(* IEC 61131-3 sources: daoli-st-library/DL_Device (part 26) *)

(* ---- FB_DL_MfcFlowCtrl.st ---- *)
(*==============================================================================
 * 组件名称 (Component)  : FB_DL_MfcFlowCtrl
 * 所属子库 (Sublibrary) : DL_Device
 * 当前版本 (Version)    : 1.0.1
 * 兼容性 (Platform)     : CODESYS 3.5 / TwinCAT 3 / 汇川 InoProShop / Machine Expert
 *                         仅依赖纯 IEC 61131-3 标准元素，零厂商方言
 * 功能描述 (Function)   : MFC 设定-回读校验：新设定上升沿启动跟踪窗，窗内峰值
 *                         对设定+超调阈判超调；回读持续 tStable 在容差窗内判
 *                         入容差；跟踪窗超时（tStable x 5）未入窗 → 稳定超时故障。
 *                         设定 0 视为关断不校验；回读 NaN/越量程判无效冻结。
 * 溯源 (Origin)         : 道莅 clean-room 防御性实现
 * 本文件内含 (Contains) : TYPE E_DL_MfcState / TYPE E_DL_MfcErr /
 *                         FUNCTION_BLOCK FB_DL_MfcFlowCtrl
 * 依赖 (Depends)        : DL_MathData/FC_DL_TimeToDintMs、DL_MathData/FC_DL_TimeScaleSat
 * 红线自检 (Redline)    : 无外部全局变量、无硬件地址直引 ｜ 全变量中英双语同行注释
 *                         防除零 + 参数下限钳制 + 非有限值防御 ｜ 枚举成员全部显式赋值
 *                         TON/沿检测实例每周期无条件调用（仅 IN 条件化）｜
 *                         跟踪窗状态机 CASE 含 ELSE 兜底 ｜ 峰值检测用比较禁浮点判等
 * 错误码表 (Codes)      : 16#0003_0398 就绪
 *                         16#0003_0399 校验通过
 *                         16#0003_039A 信息级 超调检出（不阻断判据）
 *                         16#0003_039B 故障级 稳定超时
 *                         16#0003_039C 故障级 回读无效（冻结判定）
 * 修订历史 (Revision)   : 2026-11-17  v1.0.0  首版入库 · R27 · 阶段三批 2
 *                         2026-11-17  v1.0.1  R27 终审修复（对外引脚零变更）：超调峰值改为
 *                         「首次入窗后才累积、初值取设定」。原实现 fPeakSlm 初值取当前回读，
 *                         降设定（如 20→10 slm）时回读 20 立即满足 20−10 > 超调阈，
 *                         每次下调设定必误报 039A 超调；改为入窗锁存后，仅真实向上超调计入。
 * 验收向量 (Acceptance) : 设定 10 slm 容差 2%FS 超调阈 5%FS：回读峰值 11.0 slm
 *                         → 超调 10%FS → 039A；回读持续 5 s 在 9.8~10.2 → 0399；
 *                         回读 8 slm 持续 25 s → 039B
 *============================================================================*)

(*-----------------------------------------------------------------------------
 * 枚举: E_DL_MfcState（归属 DL_Device，跟踪窗状态机状态）
 *----------------------------------------------------------------------------*)
TYPE E_DL_MfcState :
(
    eIdle    := 0,    // 就绪待新设定 / Idle, waiting for a new setpoint
    eTrack   := 10,   // 跟踪窗：峰值检测与入窗监视 / Tracking window, peak and entry watch
    eStable  := 20,   // 稳定窗：持续容差内计时 / Stable window, dwell timing
    eDone    := 30,   // 校验通过（可被新设定重开）/ Verification passed
    eTimeout := 40,   // 稳定超时故障 / Stable timeout fault
    eFault   := 99    // 回读无效兜底态 / Readback-invalid fallback
);
END_TYPE

(*-----------------------------------------------------------------------------
 * 枚举: E_DL_MfcErr（归属 DL_Device，与 FB_DL_MfcFlowCtrl 同文件）
 *----------------------------------------------------------------------------*)
TYPE E_DL_MfcErr :
(
    eReady      := 16#0003_0398,   // 就绪 / Ready
    ePass       := 16#0003_0399,   // 校验通过 / Verification passed
    eOvershoot  := 16#0003_039A,   // 信息级：超调检出 / Info: overshoot detected
    eStableTmo  := 16#0003_039B,   // 故障级：稳定超时 / Fault: stable timeout
    eReadbackBad:= 16#0003_039C    // 故障级：回读无效 / Fault: readback invalid
);
END_TYPE

(*==============================================================================
 * 功能块: FB_DL_MfcFlowCtrl
 * 调用约定: 每个扫描周期无条件调用一次；tSampleTime 注入真实任务间隔。
 *============================================================================*)
FUNCTION_BLOCK FB_DL_MfcFlowCtrl
VAR_INPUT
    fSetpointSlm   : REAL;            // 设定流量 [标准升每分钟]，有效域 0~满量程 / Setpoint flow [slm]
    fReadbackSlm   : REAL;            // 回读流量 [标准升每分钟] / Readback flow [slm]
    fScaleMaxSlm   : REAL;            // MFC 满量程 [标准升每分钟]，须 > 0 / MFC full scale [slm]
    fTolPct        : REAL := 2.0;     // 容差 [%FS]，默认 2，下限钳 0.5 / Tolerance [percent of FS]
    fOvershootPct  : REAL := 5.0;     // 超调判据 [%FS]，默认 5，下限钳 0.5 / Overshoot criterion [percent of FS]
    tStable        : TIME := T#5S;    // 稳定窗时长 [秒] / Stable window duration [s]
    bNewSp         : BOOL;            // 新设定触发（上升沿）/ New setpoint trigger, rising edge
    tSampleTime    : TIME := T#100MS; // 采样周期，调用方注入 / Sample period, caller-injected
END_VAR
VAR_OUTPUT
    bInTol         : BOOL;            // 入容差标志 / Within-tolerance flag
    bOvershoot     : BOOL;            // 超调检出标志 / Overshoot detected flag
    tSettleMs      : UDINT;           // 实测稳定时间 [毫秒] / Measured settle time [ms]
    eError         : E_DL_MfcErr;     // 错误码 / Error code
    eState         : E_DL_MfcState;   // 跟踪窗状态机当前状态 / Tracking window state
END_VAR
VAR
    fbNewSpTrig    : R_TRIG;          // 新设定上升沿实例（无条件调用）/ New setpoint edge instance
    fbTonStable    : TON;             // 稳定窗计时器（无条件调用）/ Stable window timer
    fbTonWindow    : TON;             // 跟踪窗超时计时器（无条件调用）/ Tracking window timeout timer
    fPeakSlm       : REAL;            // 跟踪窗内回读峰值 [标准升每分钟] / Readback peak in window [slm]
    fTolAbs        : REAL;            // 容差绝对值 [标准升每分钟] / Tolerance in absolute flow [slm]
    fOverAbs       : REAL;            // 超调阈绝对值 [标准升每分钟] / Overshoot threshold in absolute flow [slm]
    fSpUse         : REAL;            // 生效设定（NaN 兜底）[标准升每分钟] / Effective setpoint [slm]
    fScaleUse      : REAL;            // 生效满量程（NaN 兜底）[标准升每分钟] / Effective full scale [slm]
    bReadOk        : BOOL;            // 回读有效性判据 / Readback validity predicate
    uMsErr         : UDINT;           // 委托时间换算错误码（0 = 无错）/ Delegate time-conversion error id
    bInWin         : BOOL;            // 回读在容差窗内（瞬时）/ Readback within window, instantaneous
    bReached       : BOOL;            // 本窗内首次入窗锁存（v1.0.1：峰值仅此后计入）/ First-in-window latch, peak counted afterwards
END_VAR
VAR CONSTANT
    DL_MFC_TOL_MIN    : REAL := 0.5;     // 容差下限 [%FS] / Tolerance lower bound [percent FS]
    DL_MFC_OVER_MIN   : REAL := 0.5;     // 超调阈下限 [%FS] / Overshoot lower bound [percent FS]
    DL_MFC_PCT        : REAL := 100.0;   // 百分数系数 [百分数] / Percent factor
    DL_MFC_WINDOW_K   : INT  := 5;       // 跟踪窗超时倍率（tStable x 5）/ Tracking window timeout multiplier
    DL_MFC_INF_MAX    : REAL := 1.0E30;  // 非有限值判定幅值上限 / Magnitude bound for finite-value check
    DL_MFC_ZERO       : REAL := 0.0;     // 零值常量，避免裸字面量 / Zero constant
    DL_MFC_MS_CAP     : UDINT := 16#FFFF_FFFE;   // 稳定时间输出饱和值 [毫秒] / Settle time saturation [ms]
END_VAR

(*------------------------------------------------------------------------------
 * 段 1｜沿检测与 TON 实例每周期无条件调用（仅 IN 条件化）
 *----------------------------------------------------------------------------*)
fbNewSpTrig(CLK := bNewSp);                           // 新设定沿检测无条件刷新 / new setpoint edge refreshed unconditionally
fbTonStable(IN := (eState = E_DL_MfcState.eStable) AND bInWin, PT := tStable);        // 稳定窗计时 / stable dwell timing
fbTonWindow(IN := (eState = E_DL_MfcState.eTrack), PT := FC_DL_TimeScaleSat(tIn := tStable, nScale := DL_MFC_WINDOW_K));   // 跟踪窗超时计时（tStable x 5，委托换算）/ tracking window timing via delegate

(*------------------------------------------------------------------------------
 * 段 2｜参数防御：满量程/设定 NaN 兜底，容差与超调下限钳 0.5 %FS
 *----------------------------------------------------------------------------*)
fScaleUse := fScaleMaxSlm;                            // 满量程工作副本 / full-scale working copy
IF (fScaleUse <> fScaleUse) OR (fScaleUse <= DL_MFC_ZERO) OR (fScaleUse > DL_MFC_INF_MAX) THEN
    fScaleUse := 100.0;                               // 满量程非法按 100 slm 兜底 / illegal full scale falls back to 100 slm
END_IF
fSpUse := fSetpointSlm;                               // 设定工作副本 / setpoint working copy
IF (fSpUse <> fSpUse) OR (ABS(fSpUse) > DL_MFC_INF_MAX) THEN
    fSpUse := DL_MFC_ZERO;                            // 设定非有限按 0（关断语义）/ non-finite setpoint treated as zero
END_IF
IF fTolPct < DL_MFC_TOL_MIN THEN
    fTolAbs := fScaleUse * DL_MFC_TOL_MIN / DL_MFC_PCT;   // 容差下限钳制 [标准升每分钟] / tolerance floored [slm]
ELSIF fTolPct > DL_MFC_PCT THEN
    fTolAbs := fScaleUse;                             // 容差上限钳制（满量程封顶）/ tolerance capped at FS
ELSE
    fTolAbs := fScaleUse * fTolPct / DL_MFC_PCT;      // 容差换算 [标准升每分钟] / tolerance computed [slm]
END_IF
IF fOvershootPct < DL_MFC_OVER_MIN THEN
    fOverAbs := fScaleUse * DL_MFC_OVER_MIN / DL_MFC_PCT;   // 超调阈下限钳制 / overshoot floored
ELSIF fOvershootPct > DL_MFC_PCT THEN
    fOverAbs := fScaleUse;                            // 超调阈上限钳制 / overshoot capped at FS
ELSE
    fOverAbs := fScaleUse * fOvershootPct / DL_MFC_PCT;   // 超调阈换算 / overshoot computed
END_IF

(*------------------------------------------------------------------------------
 * 段 3｜回读有效性判据：NaN/越量程/负值判无效（bReadOk 为 FALSE 时冻结判定）
 *----------------------------------------------------------------------------*)
bReadOk := (fReadbackSlm = fReadbackSlm)                      // 自反判 NaN / NaN self-reflexive test
        AND (ABS(fReadbackSlm) <= DL_MFC_INF_MAX)             // 溢出判 / overflow test
        AND (fReadbackSlm >= DL_MFC_ZERO)                     // 负流量无效 / negative flow invalid
        AND (fReadbackSlm <= fScaleUse * 1.5);                // 越量程 150% 判无效 / over-range 150 percent invalid

(*------------------------------------------------------------------------------
 * 段 4｜瞬时入窗判据：|回读 - 设定| <= 容差（比较判据，禁浮点判等）
 *----------------------------------------------------------------------------*)
bInWin := bReadOk AND (ABS(fReadbackSlm - fSpUse) <= fTolAbs);   // 瞬时入窗 / instantaneous in-window
IF bInWin THEN
    bReached := TRUE;                                 // v1.0.1：首次入窗锁存，此后峰值才计 / latch on first entry, peak counted after
END_IF
bInTol := bInWin AND fbTonStable.Q AND (eState <> E_DL_MfcState.eIdle);   // 入容差 = 瞬时 + 持续达时 / in-tol combined

(*------------------------------------------------------------------------------
 * 段 5｜新设定上升沿：重开跟踪窗（设定 0 关断不校验，直回就绪）
 *----------------------------------------------------------------------------*)
IF fbNewSpTrig.Q THEN
    IF (fSpUse <= DL_MFC_ZERO) OR (NOT bReadOk) THEN
        eState := E_DL_MfcState.eIdle;                // 设定 0 或回读无效：不启动校验 / zero setpoint or bad readback: no verify
    ELSE
        eState := E_DL_MfcState.eTrack;               // 启动跟踪窗 / start tracking window
        fPeakSlm := fSpUse;                           // v1.0.1：峰值初值取设定而非回读 / peak preset to setpoint, not readback
        bReached := FALSE;                            // v1.0.1：首次入窗锁存清零 / first-entry latch cleared
        bOvershoot := FALSE;                          // 超调标志清零 / overshoot flag cleared
        tSettleMs := 0;                               // 稳定时间清零 / settle time cleared
    END_IF
END_IF

(*------------------------------------------------------------------------------
 * 段 6｜跟踪窗状态机：CASE 含 ELSE 兜底
 *----------------------------------------------------------------------------*)
CASE eState OF

    E_DL_MfcState.eIdle:
        bInTol := FALSE;                              // 就绪态无入容差 / no in-tol in idle
        bOvershoot := FALSE;                          // 就绪态无超调 / no overshoot in idle
        tSettleMs := 0;                               // 稳定时间清零 / settle time cleared
        eError := E_DL_MfcErr.eReady;                 // 码 0398 / code ready

    E_DL_MfcState.eTrack:
        IF bReadOk AND bReached THEN
            IF fReadbackSlm > fPeakSlm THEN
                fPeakSlm := fReadbackSlm;             // 峰值更新（仅首次入窗后计入，禁浮点判等）/ peak after first entry
            END_IF
            IF (fPeakSlm - fSpUse) > fOverAbs THEN
                bOvershoot := TRUE;                   // 超调检出 / overshoot detected
            END_IF
        END_IF
        IF NOT bReadOk THEN
            eState := E_DL_MfcState.eFault;           // 回读无效：冻结进兜底态 / readback invalid: freeze to fallback
            eError := E_DL_MfcErr.eReadbackBad;       // 故障级：回读无效 / fault: readback invalid
        ELSIF bInWin AND fbTonStable.Q THEN
            eState := E_DL_MfcState.eDone;            // 窗内已达标：直接通过（极快稳定路径）/ fast-pass path
        ELSIF bInWin THEN
            eState := E_DL_MfcState.eStable;          // 入窗：进稳定窗 / entered window: stable phase
        ELSIF fbTonWindow.Q THEN
            eState := E_DL_MfcState.eTimeout;         // 跟踪窗超时（tStable x 5）/ tracking window timeout
            eError := E_DL_MfcErr.eStableTmo;         // 故障级：稳定超时 / fault: stable timeout
        ELSE
            eError := E_DL_MfcErr.eReady;             // 跟踪中先挂就绪码 / ready code while tracking
        END_IF

    E_DL_MfcState.eStable:
        IF NOT bReadOk THEN
            eState := E_DL_MfcState.eFault;           // 回读无效：冻结进兜底态 / readback invalid: freeze
            eError := E_DL_MfcErr.eReadbackBad;       // 故障级：回读无效 / fault: readback invalid
        ELSIF fbTonStable.Q THEN
            eState := E_DL_MfcState.eDone;            // 持续在窗达 tStable：通过 / dwell met: passed
            IF bOvershoot THEN
                eError := E_DL_MfcErr.eOvershoot;     // 信息级：超调检出（通过但留痕）/ info: overshoot noted
            ELSE
                eError := E_DL_MfcErr.ePass;          // 码 0399 / code pass
            END_IF
            tSettleMs := DINT_TO_UDINT(FC_DL_TimeToDintMs(tIn := fbTonStable.ET, eErr => uMsErr));   // 实测稳定时间委托换算 [毫秒] / settle time via delegate [ms]
            IF (uMsErr <> 0) OR (tSettleMs > DL_MFC_MS_CAP) THEN
                tSettleMs := DL_MFC_MS_CAP;           // 换算失败或越界：饱和输出 / conversion failure saturates
            END_IF
        ELSIF NOT bInWin THEN
            eState := E_DL_MfcState.eTrack;           // 出窗：回跟踪窗继续监视（计时随 IN 断开自清）/ left window: back to tracking
            eError := E_DL_MfcErr.eReady;             // 回挂就绪码 / ready code again
        END_IF

    E_DL_MfcState.eDone:
        bInTol := TRUE;                               // 通过态保持入容差显示 / in-tol held on pass
        IF fbNewSpTrig.Q THEN
            eError := E_DL_MfcErr.eReady;             // 新设定沿已由段 5 处理 / new setpoint handled in section 5
        END_IF

    E_DL_MfcState.eTimeout:
        bInTol := FALSE;                              // 超时态入容差撤销 / in-tol dropped on timeout
        // 稳定超时为故障级：码 039B 已在转出时置位，保持至新设定沿 / fault code 039B held until next setpoint edge

    E_DL_MfcState.eFault:
        bInTol := FALSE;                              // 兜底态入容差撤销 / in-tol dropped
        IF NOT bReadOk THEN
            eError := E_DL_MfcErr.eReadbackBad;       // 回读仍无效：保持故障码 / readback still invalid: hold code
        ELSE
            eState := E_DL_MfcState.eIdle;            // 回读恢复：自动回就绪 / readback recovered: back to idle
            eError := E_DL_MfcErr.eReady;             // 回就绪码 / ready code
        END_IF

    ELSE
        eState := E_DL_MfcState.eFault;               // 非法状态兜底 / illegal-state fallback
        eError := E_DL_MfcErr.eReadbackBad;           // 兜底码（回读无效段，反证句：输出同为全撤+故障级）/ fallback code
        bInTol := FALSE;                              // 入容差撤 / in-tol dropped
        bOvershoot := FALSE;                          // 超调撤 / overshoot dropped

END_CASE
END_FUNCTION_BLOCK

(* ---- FB_DL_MfcRatioCheck.st ---- *)
(*
  FB_DL_MfcRatioCheck  —  MFC 流量配比偏差核对 / MFC flow ratio deviation check
  分类 Category : DL_Device
  码位 Code     : 16#03_2_02
  版本 Version  : 1.0.0
  溯源 Source   : LBP 语义借鉴 · clean-room 实现，仅借分类/参数域/命名，未复制源码
  功能 Function : 1) 各路流量经标定换算（增益/偏置）后计算配比，与配比设定窗比对；
                  2) 设定回读比对带容差（浮点禁 = 判等），差异只报等级不改设定值；
                  3) 配比计算前各路流量须 > 0 且有限（分母防零），配比窗上下限须配比校验。
  边界 Boundary : ① 配比计算前各路流量 > 0 且有限（分母防零）；
                  ② 配比窗上下限配比校验（下限 <= 上限），倒置即报码；
                  ③ 设定回读比对带容差，差异只报等级不改设定值；
                  ④ 输出三行同向：配比实测 → 配比判定 → 回读不一致标志。
  依赖 Depends  : FB_DL_DeviceParamVerify（设定回读比对，每拍无条件调用）

  码表 Error codes（本件子码步进 16#10，避让邻件码位）:
    16#0002_0302 故障级：组态非法（配比窗倒置 / 标定增益 <= 0 / 路数越界 / 容差 <= 0）
    16#0002_0312 故障级：回读参数超差（不一致锁存）
    16#0002_0322 信息级：某路流量为 0 或非有限，本拍不出配比结论（不置 bError）
*)

TYPE E_DL_MrcPhase :
(
    eIdle    := 0,   // 空闲 / Idle
    eCalc    := 10,  // 配比计算 / Ratio computation
    eVerify  := 20,  // 回读比对 / Readback verification
    eVerdict := 30,  // 结论输出 / Verdict output
    eFault   := 90   // 故障锁定 / Fault locked
);
END_TYPE

FUNCTION_BLOCK FB_DL_MfcRatioCheck
VAR_INPUT
    bEnable      : BOOL;                          // 总使能，FALSE 回空闲 / Master enable
    bSample      : BOOL := TRUE;                  // 采样使能 / Sampling enable
    bReset       : BOOL;                          // 复位，上升沿清故障与比对锁存 / Reset
    bAcknowledge : BOOL;                          // 上升沿确认回读不一致 / Rising edge acknowledges a mismatch
    nGasCount    : INT := 2;                      // 参与配比的气路数 [路]，域 2~4 / Participating gas channels, 2..4
    afFlowSccm   : ARRAY[1..4] OF REAL;           // 各路实测流量 [sccm] / Per-channel measured flow [sccm]
    afCalGain    : ARRAY[1..4] OF REAL;           // 各路标定增益 [sccm 折算比]，域 > 0 / Per-channel calibration gain
    afCalOffset  : ARRAY[1..4] OF REAL;           // 各路标定偏置 [sccm] / Per-channel calibration offset [sccm]
    fRatioSetPct : REAL := 50.0;                  // 配比设定（第 1 路占比）[%]，域 0~100 / Ratio setpoint [%]
    fRatioWinLo  : REAL := 45.0;                  // 配比窗下限 [%] / Ratio window low [%]
    fRatioWinHi  : REAL := 55.0;                  // 配比窗上限 [%] / Ratio window high [%]
    afSpCmd      : ARRAY[1..4] OF REAL;           // 各路设定指令 [sccm] / Per-channel setpoint command [sccm]
    afSpReadback : ARRAY[1..4] OF REAL;           // 各路设定回读 [sccm] / Per-channel setpoint readback [sccm]
    fReadbackTol : REAL := 1.0;                   // 回读容差 [sccm]（浮点禁 = 判等）/ Readback tolerance [sccm]
    fEps         : REAL := 1.0E-6;                // 浮点判零容差 [1] / Floating zero tolerance
END_VAR
VAR_OUTPUT
    fRatioActPct : REAL;                          // 实测配比（第 1 路占比）[%] / Measured ratio [%]
    fTotalFlow   : REAL;                          // 标定后总流量 [sccm] / Calibrated total flow [sccm]
    bRatioOk     : BOOL;                          // 配比在窗内 / Ratio inside window
    bFlowInvalid : BOOL;                          // 流量无效标志（0 或非有限）/ Flow invalid flag
    bMismatch    : BOOL;                          // 回读不一致（保持型）/ Readback mismatch, held
    nDiffCount   : INT;                           // 回读超差路数 [路] / Out-of-tolerance channel count
    bError       : BOOL;                          // 故障标志，与故障级码配对 / Fault flag paired with fault codes
    uErrorId     : UDINT;                         // 事件码，0 = 无事件 / Event code, 0 = none
    eStateOut    : E_DL_MrcPhase;                 // 状态机当前态，段尾单点映射 / Phase mapped at tail
END_VAR
VAR
    _eState      : E_DL_MrcPhase := E_DL_MrcPhase.eIdle;  // 内部状态 / Internal state
    rtrReset     : R_TRIG;                        // 复位沿 / Reset edge
    fbVerify     : FB_DL_DeviceParamVerify;       // 回读比对实例（无条件调用）/ Readback verify instance
    afExp       : ARRAY[1..64] OF REAL;           // 期望参数块（映射到前 4 项）/ Expected parameter block
    afAct       : ARRAY[1..64] OF REAL;           // 实际参数块（映射到前 4 项）/ Actual parameter block
    afTol       : ARRAY[1..64] OF REAL;           // 逐项容差块 / Per-item tolerance block
    nN           : INT;                           // 钳位后气路数 [路] / Clamped channel count
    nI           : INT;                           // 气路循环下标 / Channel loop index
    nDiff        : INT;                           // 本地超差计数 [路] / Local difference counter
    bCfgOk       : BOOL;                          // 组态合法标志 / Configuration valid
    bFlowOk      : BOOL;                          // 全部气路流量有效 / All flows valid
    fCalc        : REAL;                          // 单路标定后流量 [sccm] / Calibrated channel flow [sccm]
    fSum         : REAL;                          // 总流量累计 [sccm] / Total flow accumulator [sccm]
    fFirst       : REAL;                          // 第 1 路标定后流量 [sccm] / Channel-1 calibrated flow [sccm]
    uFault       : UDINT;                         // 锁存故障码 / Latched fault code
    uInfo        : UDINT;                         // 信息级码 / Information code
END_VAR
VAR CONSTANT
    DL_MRC_CHMAX : INT := 4;                      // 气路上界 [路] / Channel upper bound
    DL_MRC_PCTMAX: REAL := 100.0;                 // 百分比满量程 [%] / Percentage full scale
    DL_MRC_FLMAX : REAL := 1.0E5;                 // 单路流量物理域上限 [sccm] / Channel flow domain high
END_VAR

(* === 段 0 · 实例刷新（无条件周期调用）=== *)
rtrReset(CLK := bReset);                          // 每拍刷新复位沿

(* === 段 1 · 组态闸 === *)
nN := nGasCount;                                  // 气路数取用前钳位
IF nN < 2 THEN
    nN := 2;                                      // 配比至少两路
END_IF
IF nN > DL_MRC_CHMAX THEN
    nN := DL_MRC_CHMAX;                           // 上限钳位
END_IF
bCfgOk := (nGasCount >= 2) AND (nGasCount <= DL_MRC_CHMAX)
          AND (fRatioWinHi >= fRatioWinLo)                              // 配比窗配比校验（下限 <= 上限）
          AND (fRatioWinLo >= 0.0) AND (fRatioWinHi <= DL_MRC_PCTMAX)
          AND (fReadbackTol > fEps) AND (fRatioSetPct = fRatioSetPct)
          AND (fRatioWinLo = fRatioWinLo) AND (fRatioWinHi = fRatioWinHi);   // 含 NaN 自反
FOR nI := 1 TO DL_MRC_CHMAX DO
    IF nI <= nN THEN
        bCfgOk := bCfgOk AND (afCalGain[nI] > fEps)                    // 标定增益正域（防换算除零/反向）
                  AND (afCalGain[nI] = afCalGain[nI])                  // 增益 NaN 自反
                  AND (afCalOffset[nI] = afCalOffset[nI]);             // 偏置 NaN 自反
    END_IF
END_FOR
IF NOT bCfgOk THEN
    uFault := 16#0002_0302;                       // 故障级：组态非法
END_IF
IF rtrReset.Q AND bCfgOk THEN
    uFault := 16#0000;                            // 复位沿清锁存（复位路径可达）
    bMismatch := FALSE;                           // 回读不一致同步复位
END_IF
uInfo := 16#0000;                                 // 信息码每拍清零

(* === 段 2 · 标定换算与流量有效域（分母防零前置）=== *)
bFlowOk := TRUE;                                  // 假定有效，逐路否决
fSum := 0.0;                                      // 总流量清零
fFirst := 0.0;                                    // 第 1 路清零
FOR nI := 1 TO DL_MRC_CHMAX DO
    IF nI <= nN THEN
        IF (afFlowSccm[nI] = afFlowSccm[nI]) AND (ABS(afFlowSccm[nI]) < 1.0E30)
           AND (afFlowSccm[nI] > 0.0) AND (afFlowSccm[nI] <= DL_MRC_FLMAX) THEN
            fCalc := afFlowSccm[nI] * afCalGain[nI] + afCalOffset[nI];   // 标定换算
            IF fCalc < 0.0 THEN
                fCalc := 0.0;                                          // 负流量截零（物理不可达）
            END_IF
            fSum := fSum + fCalc;                                      // 总流量累加
            IF nI = 1 THEN
                fFirst := fCalc;                                       // 第 1 路流量
            END_IF
        ELSE
            bFlowOk := FALSE;                                          // 该路无效：本拍不出配比结论
        END_IF
    END_IF
END_FOR
bFlowInvalid := NOT bFlowOk;                      // 流量无效标志

(* === 段 3 · 比对参数块装配 + 比对实例无条件调用（先刷新，后判定）=== *)
FOR nI := 1 TO DL_MRC_CHMAX DO
    IF nI <= nN THEN
        afExp[nI] := afSpCmd[nI];                 // 期望参数装入（前 nN 项）
        afAct[nI] := afSpReadback[nI];            // 实际参数装入
        afTol[nI] := fReadbackTol;                // 逐项容差
    ELSE
        afExp[nI] := 0.0;                         // 未用项置 0（比对块按 nN 取项）
        afAct[nI] := 0.0;                         // 未用项置 0
        afTol[nI] := fReadbackTol;                // 未用项容差给默认，不影响 nN 内比对
    END_IF
END_FOR
fbVerify(bEnable := bEnable AND bCfgOk,           // 组态非法不比对
         bReset := rtrReset.Q,                    // 复位沿清比对锁存
         bAcknowledge := bAcknowledge,            // 人工确认不一致
         nItemCount := nN,                        // 比对项数 = 气路数（已钳位 2..4）
         afExpected := afExp,                     // 期望参数块
         afActual := afAct,                       // 回读参数块
         afTolerance := afTol,                    // 逐项容差（浮点禁 = 判等）
         fDefaultTol := fReadbackTol,             // 默认容差
         tVerifyTimeout := T#5S);                 // 回读超时 [ms]

(* === 段 4 · 主状态机（ENUM + CASE，含 ELSE 兜底）=== *)
CASE _eState OF
E_DL_MrcPhase.eIdle :
    bRatioOk := FALSE;                            // 空闲无配比结论
    nDiffCount := 0;                              // 超差路数清零
    IF uFault = 16#0002_0302 THEN
        _eState := E_DL_MrcPhase.eFault;          // 组态故障优先
    ELSIF bEnable AND bSample THEN
        _eState := E_DL_MrcPhase.eCalc;           // 进入计算相
    END_IF

E_DL_MrcPhase.eCalc :
    IF (NOT bFlowOk) OR (NOT bCfgOk) THEN
        bRatioOk := FALSE;                        // 无效：不出配比结论
        uInfo := 16#0002_0322;                    // 信息级：某路流量无效
    ELSIF fSum > fEps THEN
        fTotalFlow := fSum;                       // 总流量输出
        fRatioActPct := fFirst / fSum * DL_MRC_PCTMAX;   // 配比 = 第 1 路 / 总流量，分母已判非零
        bRatioOk := (fRatioActPct >= fRatioWinLo - fEps) AND (fRatioActPct <= fRatioWinHi + fEps);  // 容差窗比对
    ELSE
        fTotalFlow := 0.0;                        // 总流量近零：配比不可算
        bRatioOk := FALSE;                        // 不给结论（防除零）
        uInfo := 16#0002_0322;                    // 信息级：总流量近零
    END_IF
    _eState := E_DL_MrcPhase.eVerify;             // 转回读比对相

E_DL_MrcPhase.eVerify :
    nDiff := fbVerify.nDiffCount;                 // 取实例超差项数（本拍已刷新）
    _eState := E_DL_MrcPhase.eVerdict;            // 转结论相

E_DL_MrcPhase.eVerdict :
    nDiffCount := fbVerify.nDiffCount;            // 超差路数输出
    IF fbVerify.bMismatch THEN
        bMismatch := TRUE;                        // 置位型：回读不一致（段尾不清零）
        uFault := 16#0002_0312;                   // 故障级：回读超差
    END_IF
    IF (NOT bEnable) OR rtrReset.Q THEN
        _eState := E_DL_MrcPhase.eIdle;           // 失能/复位回空闲
    ELSIF bSample THEN
        _eState := E_DL_MrcPhase.eCalc;           // 连续采样
    END_IF

E_DL_MrcPhase.eFault :
    bRatioOk := FALSE;                            // 故障态不给配比合格结论
    IF uFault = 16#0000 THEN
        _eState := E_DL_MrcPhase.eIdle;           // 解锁回空闲
    END_IF

ELSE
    _eState := E_DL_MrcPhase.eFault;              // 非法状态拦截
    uFault := 16#0002_0302;                       // 故障级：相 ID 越界
    bRatioOk := FALSE;                            // 安全侧不给合格结论
END_CASE

(* === 段 5 · 输出映射（三行同向：配比 → 判定 → 不一致标志）=== *)
IF bFlowInvalid THEN
    bRatioOk := FALSE;                            // 流量无效绝不判合格
END_IF
IF NOT bEnable THEN
    bRatioOk := FALSE;                            // 失能不给合格结论
END_IF
bError := (uFault <> 16#0000);                    // 故障标志仅由故障级码置位（R45 配对）
IF bError THEN
    uErrorId := uFault;                           // 故障级优先上报
ELSE
    uErrorId := uInfo;                            // 否则上报信息级码
END_IF
eStateOut := _eState;                             // 输出枚举段尾单点映射（N2 规则）
END_FUNCTION_BLOCK

(* ---- FB_DL_MfcSetpointRamp.st ---- *)
//==============================================================================
// 功能块：FB_DL_MfcSetpointRamp ｜ 中文名称：MFC 设定值斜坡与超调抑制
// 所属子库：DL_Device ｜ 版本：v1.0.0 ｜ 兼容：CODESYS V3.5+ / TwinCAT 3 / 汇川 InoProShop
// 功能描述：质量流量控制器（MFC）设定值斜坡——目标值先钳量程域
//           [0, fRangeSccm]，再按恒定斜率 fSlewRateSccmS 向目标逼近
//           （每拍步进 = 斜率 x 扫描周期秒），到达即锁存 bRampDone 并
//           同步输出占量程百分比设定（fSpPctOut，模拟量给定位）。bHold
//           冻结当前值（保持，不回零）。斜坡中组态漂移（量程/斜率/周期
//           变非法）→ 冻结当前值安全侧并报故障。斜率限制即超调抑制的
//           上游手段（阶跃目标被强制线性化，下游 PID 不再追大阶跃）。
// 遗留假设（R95 代理阈值三句）：① 代理值 = fCycleTimeS 组态扫描周期
//           [秒]；② 覆盖 0.001~0.1 秒（1~100 ms）任务周期范围；③
//           覆盖不到的区间（更长周期或变周期任务）由调用方按实际任务
//           周期重设 fCycleTimeS 引脚负责，该假设挂编译验证债。
// 开源溯源 (Origin)：道莅原创实现（参考 MFC 流量控制与斜坡设定工程惯例 分类与参数域）
// 单位表：设定值[标准毫升每分钟 sccm] / 量程[sccm] / 斜率[sccm每秒] /
//         扫描周期[秒] / 百分比[%] / 时间[ms]
// 错误码表：16#0003_018E 信息级（斜坡完成：目标到达，不置 bError）/
//           16#0003_018F 信息级（目标超量程已钳位照算，不置 bError）/
//           16#0003_0366 故障级（组态非法：量程/斜率/周期 <= 0 或任一
//           输入非有限，置 bError）/ 16#0003_0367 故障级（斜坡中组态
//           漂移：运行态参数变非法，冻结当前值安全侧，置 bError——
//           该场景不可由 0366 的「触发前组态」路径观测，属运行中漂移
//           独立域）/ 16#0003_0368 故障级兜底（状态机落 ELSE，置
//           bError）
// 状态机：E_DL_MfcRampState（四态：eIdle=0 / eRamping=10 / eDone=20 /
//           eFault=99），CASE 含 ELSE 兜底，ELSE 置 0368 并冻结输出
// 边界行为：① 触发前组态非法 → 故障态锁存，bReset 复位；② 目标超
//           [0, 量程] → 双侧钳位照算 + 信息 018F；③ 斜坡中 bHold →
//           冻结当前值（保持非清零），撤销后续走；④ 到达锁存：目标
//           变更须新触发沿才重启斜坡（防每拍抖动重启）；⑤ 斜坡中
//           组态漂移 → 冻结当前值 + 故障 0367；⑥ 安全侧 = 故障态
//           fSpRampedSccm 冻结为进入故障前的最后合法值，禁止跳变
//           到 0 冲击工艺腔（MFC 设定跳变比保持更危险）。
// 修订历史：v1.0.0 2026-11-17 首版（R24 派单 · ROADMAP P2 §710）
//==============================================================================

(*------------------------------------------------------------------------------
 * 枚举: E_DL_MfcRampState（归属本功能块，同文件发布，全库唯一定义）
 * 含义: 斜坡相位，每个成员在 CASE 中有且仅有一个标签。
 *-----------------------------------------------------------------------------*)
TYPE E_DL_MfcRampState :
(
    eIdle    := 0,   // 空闲：等触发沿 / Idle, awaiting trigger edge
    eRamping := 10,  // 斜坡中：恒斜率逼近目标 / Ramping, constant slew toward the target
    eDone    := 20,  // 完成：目标到达锁存 / Done, arrival latched
    eFault   := 99   // 故障：组态非法/漂移/非法状态 / Fault, config, drift or illegal state
);
END_TYPE

FUNCTION_BLOCK FB_DL_MfcSetpointRamp
VAR_INPUT
    bExecute      : BOOL;                   // 触发斜坡 [—]，上升沿生效 / Trigger the ramp, rising edge
    bHold         : BOOL;                   // 冻结保持 [—]，电平生效 / Freeze hold, level effective
    bReset        : BOOL;                   // 故障复位 [—]，上升沿清故障态 / Fault reset, rising edge clears the fault state
    fSpTargetSccm : LREAL;                  // 目标设定值 [标准毫升每分钟]，域外钳量程照算 / Target setpoint [sccm], clamped to the range
    fRangeSccm    : LREAL := 100.0;         // MFC 量程 [标准毫升每分钟]，须 > 0 / MFC full range [sccm], must be > 0
    fSlewRateSccmS: LREAL := 10.0;          // 斜率 [标准毫升每分钟每秒]，须 > 0 / Slew rate [sccm per second], must be > 0
    fCycleTimeS   : LREAL := 0.01;          // 任务扫描周期 [秒]，须 > 0（R95 代理阈值） / Task scan cycle [s], must be > 0, R95 proxy
END_VAR
VAR_OUTPUT
    fSpRampedSccm : LREAL;                  // 斜坡后设定值 [标准毫升每分钟] / Ramped setpoint [sccm]
    fSpPctOut     : LREAL;                  // 占量程百分比 [百分数]，0..100 / Percent of range [percent], 0..100
    bRampDone     : BOOL;                   // 斜坡完成 [—]（到达态电平） / Ramp done, arrival level
    eState        : E_DL_MfcRampState;      // 相位出口 [—] / Phase outlet
    eErr          : UDINT;                  // 错误码，0 = 无错，码位 16#0003_018E 起信息级、16#0003_0366 起故障级（分带见错误码表） / Error code, 0 = no error, band info/fault per the code table
    bError        : BOOL;                   // 故障级标志，仅故障级错误置位 / Fault-class flag, set only on fault-level codes
    bValid        : BOOL;                   // 输出可用标志 / Outputs usable flag
END_VAR
VAR
    fbTrig    : R_TRIG;                     // 触发沿检测（待机/完成分支同样无条件刷新） / Trigger edge detector, refreshed unconditionally
    _eState   : E_DL_MfcRampState := E_DL_MfcRampState.eIdle; // 当前相位 / Current phase
    _bCfgBad  : BOOL;                       // 触发前组态非法锁存 / Pre-trigger config fault latch
    _bDriftBad: BOOL;                       // 运行中组态漂移锁存 / In-run config drift latch
    _bInfoClamp: BOOL;                      // 目标钳位信息当拍标志 / Target-clamp info flag of this scan
    _bInfoDone: BOOL;                       // 完成信息当拍标志 / Done info flag of this scan
    _fTarget  : LREAL;                      // 生效目标（已钳量程）[标准毫升每分钟] / Effective target, clamped [sccm]
    _fStep    : LREAL;                      // 本拍步进量 [标准毫升每分钟] / Per-scan step [sccm]
    _bIllegal : BOOL;                       // 非法状态标志 / Illegal state flag
    _bInit    : BOOL := FALSE;              // 首扫标志，初值 FALSE 取非判定 / First-scan flag, tested negated
END_VAR
VAR CONSTANT
    DL_MSR_INF    : LREAL := 1.7976931348623157E308; // LREAL 幅值上限 / LREAL magnitude ceiling
    DL_MSR_EPS    : LREAL := 1.0E-6;        // 浮点判零/到达容差 [标准毫升每分钟] / Zero and arrival tolerance [sccm]
    DL_MSR_ZERO   : LREAL := 0.0;           // 零值常量，避免裸字面量 [混合] / Zero constant, avoids a bare literal
    DL_MSR_PCT    : LREAL := 100.0;         // 百分比满量程 [百分数] / Full scale percent
END_VAR

(*------------------------------------------------------------------------------
 * 段 1｜每拍预置：输出保持语义的标志预清（设定值不在预置段清零，
 *       故障态须冻结而非清零——MFC 设定跳变比保持更危险）
 *      Flags pre-cleared, setpoint deliberately not cleared here
 *-----------------------------------------------------------------------------*)
fSpPctOut  := DL_MSR_ZERO;               // 百分比先清（段 5 重算） / Percent cleared first
eErr   := 16#0000_0000;                  // 错误码每拍重算 / Error code recomputed
bError := FALSE;                         // 故障标志每拍重算 / Fault flag recomputed
bValid := FALSE;                         // 可用标志每拍重算 / Usable flag recomputed
bRampDone := FALSE;                      // 完成电平先清（段 5 重置） / Done level cleared first
_bInfoClamp := FALSE;                    // 钳位信息预清零 / Clamp info pre-cleared
_bInfoDone  := FALSE;                    // 完成信息预清零 / Done info pre-cleared
_bIllegal   := FALSE;                    // 非法状态预清零 / Illegal flag pre-cleared

(*------------------------------------------------------------------------------
 * 段 2｜首扫初始化
 *      First-scan initialisation
 *-----------------------------------------------------------------------------*)
IF NOT _bInit THEN
    _eState  := E_DL_MfcRampState.eIdle; // 相位空闲起步 / Phase starts idle
    _bCfgBad := FALSE;                   // 组态锁存清零 / Config latch cleared
    fSpRampedSccm := DL_MSR_ZERO;        // 设定值从零起步 / Setpoint starts at zero
    _bInit  := TRUE;                     // 首扫只做一次 / The first scan runs once
END_IF

(*------------------------------------------------------------------------------
 * 段 3｜触发沿无条件刷新（R40：CASE 之外每拍必调）
 *      Trigger edge refreshed unconditionally per R40
 *-----------------------------------------------------------------------------*)
fbTrig(CLK := bExecute);                 // 触发沿检测 / Trigger edge detection

(*------------------------------------------------------------------------------
 * 段 4｜组态防御闸：非有限（R79）+ 量程/斜率/周期域
 *      Configuration defense gates
 *-----------------------------------------------------------------------------*)
IF (fSpTargetSccm <> fSpTargetSccm) OR (ABS(fSpTargetSccm) > DL_MSR_INF)
   OR (fRangeSccm <> fRangeSccm) OR (ABS(fRangeSccm) > DL_MSR_INF)
   OR (fSlewRateSccmS <> fSlewRateSccmS) OR (ABS(fSlewRateSccmS) > DL_MSR_INF)
   OR (fCycleTimeS <> fCycleTimeS) OR (ABS(fCycleTimeS) > DL_MSR_INF) THEN
    _bCfgBad := TRUE;                    // 非有限归组态非法锁存 / Non-finite folded into the config latch
END_IF
IF (NOT _bCfgBad) AND ((fRangeSccm <= DL_MSR_EPS) OR (fSlewRateSccmS <= DL_MSR_EPS)
   OR (fCycleTimeS <= DL_MSR_EPS)) THEN
    _bCfgBad := TRUE;                    // 量程/斜率/周期域非法锁存 / Range, slew and cycle domains latched
END_IF

(*------------------------------------------------------------------------------
 * 段 5｜相位机（CASE 含 ELSE 兜底；状态改写只出现在分支判据内，R39）
 *      Phase machine with ELSE fallback
 *-----------------------------------------------------------------------------*)
CASE _eState OF

    E_DL_MfcRampState.eIdle:               // 空闲：触发沿且组态合法进斜坡
        IF fbTrig.Q AND (NOT _bCfgBad) THEN
            _fTarget := MIN(MAX(fSpTargetSccm, DL_MSR_ZERO), fRangeSccm); // 目标钳量程域 / Target clamped to the range
            IF ABS(_fTarget - fSpTargetSccm) > DL_MSR_EPS THEN
                _bInfoClamp := TRUE;       // 目标超量程钳位提示（信息级） / Target clamped, info
            END_IF
            _eState := E_DL_MfcRampState.eRamping; // 进斜坡 / To ramping
        ELSIF fbTrig.Q AND _bCfgBad THEN
            _eState := E_DL_MfcRampState.eFault; // 组态非法进故障 / Illegal config to fault
        END_IF

    E_DL_MfcRampState.eRamping:            // 斜坡：恒斜率逼近；bHold 冻结；漂移落故障
        // 拍 N 进入（触发沿）/ 本拍行为：步进 = 斜率 x 周期，向目标逼近 / 拍 N+1 转出：到达进 eDone
        IF _bCfgBad THEN
            _bDriftBad := TRUE;            // 运行中组态漂移锁存（冻结当前值） / In-run drift latched, value frozen
            _eState := E_DL_MfcRampState.eFault; // 进故障 / To fault
        ELSIF bHold THEN
            fSpRampedSccm := fSpRampedSccm; // 冻结保持：本拍不动（显式自持） / Hold, no movement this scan (explicit self-hold)
        ELSE
            _fStep := fSlewRateSccmS * fCycleTimeS; // 本拍步进量 [sccm] / Per-scan step
            IF fSpRampedSccm < (_fTarget - DL_MSR_EPS) THEN
                fSpRampedSccm := MIN(fSpRampedSccm + _fStep, _fTarget); // 上行逼近（饱和于目标） / Upward approach, saturated at the target
            ELSIF fSpRampedSccm > (_fTarget + DL_MSR_EPS) THEN
                fSpRampedSccm := MAX(fSpRampedSccm - _fStep, _fTarget); // 下行逼近（饱和于目标） / Downward approach, saturated at the target
            ELSE
                _bInfoDone := TRUE;        // 目标到达（信息级，拍 N 进入） / Target reached, info
                _eState := E_DL_MfcRampState.eDone; // 拍 N+1 转出：进完成锁存 / To done, latched
            END_IF
        END_IF

    E_DL_MfcRampState.eDone:               // 完成：锁存保持，新沿才重算
        IF _bCfgBad THEN
            _bDriftBad := TRUE;            // 完成态组态漂移同域锁存 / Drift latched in done
            _eState := E_DL_MfcRampState.eFault; // 进故障 / To fault
        ELSIF fbTrig.Q THEN
            _fTarget := MIN(MAX(fSpTargetSccm, DL_MSR_ZERO), fRangeSccm); // 新目标钳量程 / New target clamped
            IF ABS(_fTarget - fSpTargetSccm) > DL_MSR_EPS THEN
                _bInfoClamp := TRUE;       // 新目标钳位提示 / New target clamped, info
            END_IF
            _eState := E_DL_MfcRampState.eRamping; // 新沿重斜坡 / New edge re-ramps
        END_IF

    E_DL_MfcRampState.eFault:              // 故障：复位沿且组态恢复回空闲（设定值保持冻结值）
        IF bReset AND (NOT _bCfgBad) AND (NOT _bDriftBad) THEN
            _bDriftBad := FALSE;           // 复位清漂移锁存 / Reset clears the drift latch
            _eState := E_DL_MfcRampState.eIdle; // 回空闲（冻结值保持） / Back to idle, frozen value held
        END_IF

    ELSE                                   // 非法状态兜底（R21：CASE 必带 ELSE）
        _bIllegal := TRUE;                 // 标记非法状态 / Flag the illegal state
        _eState   := E_DL_MfcRampState.eFault; // 回故障态（设定值冻结） / Back to fault, value frozen
END_CASE

(*------------------------------------------------------------------------------
 * 段 6｜输出换算与码位出口（故障级码 3 行内置 bError，R45/R101 配对）
 *      Output scaling and code outlet, fault codes paired with bError
 *-----------------------------------------------------------------------------*)
IF ABS(fRangeSccm) > DL_MSR_EPS THEN
    fSpPctOut := MIN(MAX(fSpRampedSccm / fRangeSccm, DL_MSR_ZERO), 1.0) * DL_MSR_PCT; // 占量程百分比 [百分数]，分母已闸 / Percent of range, denominator gated
ELSE
    fSpPctOut := DL_MSR_ZERO;              // 量程退化兜底（组态闸已挡，防御路径） / Degenerate range fallback
END_IF
fSpRampedSccm := MIN(MAX(fSpRampedSccm, DL_MSR_ZERO), fRangeSccm); // 输出终值钳量程域 / Final setpoint clamped to the range
bRampDone := (_eState = E_DL_MfcRampState.eDone); // 完成电平挂状态量（R99） / Done level bound to the state

IF _bIllegal THEN
    eErr   := 16#0003_0368;                // 故障级：状态机兜底 / Fault: state machine fallback
    bError := TRUE;                        // 置故障标志 / Raise the fault flag
ELSIF _bDriftBad THEN
    eErr   := 16#0003_0367;                // 故障级：斜坡中组态漂移（冻结安全侧） / Fault: in-run config drift, frozen safe side
    bError := TRUE;                        // 置故障标志 / Raise the fault flag
ELSIF _bCfgBad THEN
    eErr   := 16#0003_0366;                // 故障级：组态非法 / Fault: illegal configuration
    bError := TRUE;                        // 置故障标志 / Raise the fault flag
ELSIF _bInfoClamp THEN
    eErr := 16#0003_018F;                  // 信息级：目标超量程已钳位 / Info: target clamped to the range
ELSIF _bInfoDone THEN
    eErr := 16#0003_018E;                  // 信息级：斜坡完成 / Info: ramp done
END_IF

bValid := (NOT bError) AND (_eState <> E_DL_MfcRampState.eIdle); // 空闲/故障输出不可用 / Outputs unusable in idle or fault
eState := _eState;                       // 相位出口 / Phase outlet
END_FUNCTION_BLOCK

(* ---- FB_DL_MotorHealthAoi.st ---- *)
(*==============================================================================
 * 组件名称 (Component)  : FB_DL_MotorHealthAoi
 * 所属子库 (Sublibrary) : DL_Device
 * 当前版本 (Version)    : 1.0.0
 * 兼容性   (Platform)   : CODESYS 3.5 / TwinCAT 3 / 汇川 InoProShop / Machine Expert
 *                         仅依赖 Standard.library（TON / R_TRIG），零厂商方言
 * 来源标签 (Source)     : rockwell-aoi（T2-6 设备级粒度族：阀 / 电机 / 夹爪之电机）
 * 功能描述 (Function)   : 电机 AOI 三分类诊断：过温 / 过载 / 启停频繁三判据各自带
 *                         独立确认延时，任一类确认即置独立锁存与独立码位（R190 归因
 *                         唯一），并给出 NE107 健康出口与停机请求；三类锁存互不覆盖。
 * 分工互引 (Boundary)   : 过温保护动作归 FB_DL_MotorPtcThermistProtect（硬保护），
 *                         健康聚合归 FB_DL_DeviceHealthArbiter；本件只做**分类诊断
 *                         与确认计时**，不替代硬保护回路，也不做多设备聚合。
 * 边界与语义披露 (Boundary disclosure) :
 *   1) 三条判据的确认延时各自独立（tTempConfirm / tOverloadConfirm / tFreqConfirm），
 *      三计时器每拍无条件刷新（红线 R7），门控挂状态量与判据量而非单拍标志（R99）。
 *   2) 过载判据用电流比值（fCurrent / fRatedCurrent），除子由组态闸保证 > 0；
 *      比值达 fOverloadRatio 且持续确认窗即确认。
 *   3) 启停频繁判据用滚动窗计数：窗口窗长 tFreqWindow（TON 自复位 R188），
 *      窗内启动沿计数达 nStartLim 且持续 tFreqConfirm 即确认。
 *   4) 非有限输入（温度 / 电流 / 额定电流）不参与判据，只保持上一拍的确认状态，
 *      并由组态闸之外的信号闸置信息级码（不锁存，不因一扫 NaN 让诊断永久失效）。
 *   5) 健康出口口径：任一锁存 -> eFailure；任一确认中 -> eMaintenanceReq；
 *      未使能 -> eUnknown；其余 eOk。出口取最严，禁按图改序。
 * 故障码表 (Error codes) :
 *   16#0003_0532 [故障级] 组态非法（阈值域 / 确认窗 / 额定电流），诊断置挂起
 *                 反证：挂起与「设备恰好在容差内」输出组合相同，无码不可区分。
 *   16#0003_0533 [故障级] 过温确认（绕组温度持续超阈），锁存至复位沿 + 温度回落
 *                 反证：三类锁存若共用码则某类永不赋值（R190），且过温与过载的
 *                 处置完全不同（通风 vs 减载），必须独立码位。
 *   16#0003_0534 [故障级] 过载确认（电流比值持续超限），锁存至复位沿 + 电流回落
 *                 反证：与过温同状态出口，仅码位可归因（R190）。
 *   16#0003_0535 [故障级] 启停频繁确认（滚动窗启动次数超限），锁存至复位沿 + 窗刷新
 *                 反证：启停频繁不停机也可能无任何其它输出变化，无码不可观测。
 * 码位总账 (Code ledger) : 16#0003_0532 / 0533 / 0534 / 0535 用
 * 归属声明 (Ownership)  : E_DL_Ne107Status 归属 DL_Device\I_DL_DeviceHealth.st，
 *                         本件只引用不重声明
 * 依赖     (Depends)    : 无 DL_ 内部依赖；Standard.library: TON / R_TRIG
 * 红线自检 (Redline)    : R1 ✓ 零全局变量 ｜ R2 ✓ 零 %I/%Q ｜ R3 ✓ 纯 IEC 61131-3
 *                         R4 ✓ 除子由组态闸保证 / 非有限三判 / 域闸全枚举
 *                         R5 ✓ 全变量双语同行注释 ｜ R6 ✓ 四态 ENUM + ELSE 兜底
 *                         R7 ✓ 四沿四计时主体最前部无条件刷新
 * 修订历史 (Revision)   : 2026-11-22  v1.0.0  首版入库（R69 构建轮 · 批 2 · N4）
 *============================================================================*)

(*-----------------------------------------------------------------------------
 * 枚举: E_DL_MotorAoiState（归属 DL_Device，与 FB_DL_MotorHealthAoi 同文件）
 *----------------------------------------------------------------------------*)
TYPE E_DL_MotorAoiState :
(
    eIdle   := 0,     // 未使能：诊断挂起 / Disabled, diagnosis suspended
    eMonitor := 10,   // 监视中：三判据确认计时 / Monitoring, three confirm timers running
    eTripped := 20,   // 已确认停机（至少一类锁存）/ Tripped, at least one cause latched
    eFault  := 99     // 组态非法：诊断拒绝 / Config illegal, diagnosis refused
);
END_TYPE

(*==============================================================================
 * 功能块: FB_DL_MotorHealthAoi
 * 调用约定: 每个扫描周期无条件调用一次。
 *============================================================================*)
FUNCTION_BLOCK FB_DL_MotorHealthAoi
VAR_INPUT
    fWindingTemp   : REAL;                 // 绕组温度 [°C] / winding temperature [°C]
    fTempLim       : REAL := 130.0;        // 过温阈 [°C]，<= 0 组态非法 / over-temperature threshold [°C]
    fCurrent       : REAL;                 // 电机电流 [A] / motor current [A]
    fRatedCurrent  : REAL := 10.0;         // 额定电流 [A]，<= 0 组态非法（除子）/ rated current [A], the divisor
    fOverloadRatio : REAL := 1.15;         // 过载比值阈 [倍]，<= 1 组态非法 / overload ratio [x]
    bStartPulse    : BOOL;                 // 启动命令（上升沿计数）/ start command, rising edge counted
    nStartLim      : INT := 6;             // 滚动窗启动次数上限 [次]，域 1..100 / start ceiling per window [times]
    tTempConfirm   : TIME := T#3S;         // 过温确认窗 [s] / over-temperature confirm window [s]
    tOverloadConfirm : TIME := T#2S;       // 过载确认窗 [s] / overload confirm window [s]
    tFreqConfirm   : TIME := T#1S;         // 启停频繁确认窗 [s] / frequent-start confirm window [s]
    tFreqWindow    : TIME := T#60S;        // 启动计数滚动窗长 [s] / rolling start-count window [s]
    bEnable        : BOOL := TRUE;         // 使能 / enable
    bReset         : BOOL;                 // 上升沿：清三类锁存（须对应判据已消）/ rising edge clears the three latches
END_VAR
VAR_OUTPUT
    eHealth        : E_DL_Ne107Status;     // NE107 健康出口（六态，属主 I_DL_DeviceHealth）/ NE107 health verdict
    bTripReq       : BOOL;                 // 停机请求（任一锁存即 TRUE）/ stop request, any latch
    bOverTemp      : BOOL;                 // 过温锁存 / over-temperature latched
    bOverload      : BOOL;                 // 过载锁存 / overload latched
    bFreqStart     : BOOL;                 // 启停频繁锁存 / frequent-start latched
    bError         : BOOL;                 // 故障标志（组态 / 三类锁存归并）/ fault flag
    uErrorId       : UDINT;                // 故障码，0 = 无故障 / error code, 0 = none
    eState         : E_DL_MotorAoiState;   // 当前状态（供 HMI 诊断）/ current state
END_VAR
VAR
    fbTrigReset    : R_TRIG;               // 复位沿检测实例 / reset edge detector
    fbTrigStart    : R_TRIG;               // 启动命令沿检测实例 / start command edge detector
    tonTemp        : TON;                  // 过温确认计时实例 / over-temperature confirm timer
    tonOverload    : TON;                  // 过载确认计时实例 / overload confirm timer
    tonFreq        : TON;                  // 启停频繁确认计时实例 / frequent-start confirm timer
    tonFreqWin     : TON;                  // 启动计数滚动窗（自复位 R188）/ rolling window timer, self resetting
    eStateInt      : E_DL_MotorAoiState;   // 主状态机内部当前态 / internal state
    bTempCond      : BOOL;                 // 本拍过温判据成立 / over-temperature criterion true this scan
    bOvldCond      : BOOL;                 // 本拍过载判据成立 / overload criterion true this scan
    bFreqCond      : BOOL;                 // 本拍启停频繁判据成立 / frequent-start criterion true this scan
    fCurrentRatio  : REAL;                 // 电流比值 [倍]（除子已由组态闸保证 > 0）/ current ratio [x]
    nStartCnt      : INT;                  // 滚动窗内启动次数 [次] / starts inside the rolling window
    bTempLatch     : BOOL;                 // 过温锁存内部副本 / internal over-temperature latch
    bOvldLatch     : BOOL;                 // 过载锁存内部副本 / internal overload latch
    bFreqLatch     : BOOL;                 // 启停频繁锁存内部副本 / internal frequent-start latch
    bSigBad        : BOOL;                 // 温度 / 电流信号非有限 / temperature or current non-finite
    bCfgBad        : BOOL;                 // 本拍组态非法 / config illegal this scan
    bCfgLatch      : BOOL;                 // 组态锁存（复位沿 + 组态改对解除）/ config latch
    bErrorInt      : BOOL;                 // 本拍故障置位累加 / fault set accumulator
    bFirstScan     : BOOL := TRUE;         // 上电首扫标志 / first-scan flag
END_VAR
VAR CONSTANT
    DL_MH_FIN_LIM  : REAL := 1.0E30;       // REAL 幅值兜底判界 / REAL magnitude bound
    DL_MH_START_MAX : INT := 100;          // 启动次数上限闸 [次]（防计数溢出）/ start count ceiling
    DL_MH_RATIO_MIN : REAL := 1.0;         // 过载比值下限 [倍]（< 1 即常真）/ overload ratio floor [x]
END_VAR

(*------------------------------------------------------------------------------
 * 段 1｜无条件刷新区（红线 R7）：二沿四计时全部位于主体最前部
 *      Unconditional refresh: two edges and four timers at the very top
 *-----------------------------------------------------------------------------*)
fbTrigReset(CLK := bReset);
fbTrigStart(CLK := bStartPulse);
tonFreqWin(IN := NOT tonFreqWin.Q, PT := tFreqWindow);   // 自复位滚动窗（R188）/ self-resetting window

(* 段 2｜每拍预清（FB32-1）：单拍标志，禁入锁存 / per-scan preset *)
bErrorInt := FALSE;

(* 段 3｜上电首扫：三类锁存与计数落安全侧 / first-scan init *)
IF bFirstScan THEN
    eStateInt := E_DL_MotorAoiState.eIdle;
    bTempLatch := FALSE;
    bOvldLatch := FALSE;
    bFreqLatch := FALSE;
    nStartCnt  := 0;
    bFirstScan := FALSE;
END_IF

(*------------------------------------------------------------------------------
 * 段 4｜组态域闸（R151 全枚举）+ 解除路径（R152 自证可达）
 *      Config gate over every threshold, window and divisor, with the clear path
 *-----------------------------------------------------------------------------*)
bCfgBad := (fTempLim <= 0.0) OR (fTempLim <> fTempLim)
           OR (fRatedCurrent <= 0.0) OR (fRatedCurrent <> fRatedCurrent)
           OR (fOverloadRatio <= DL_MH_RATIO_MIN) OR (fOverloadRatio <> fOverloadRatio)
           OR (nStartLim < 1) OR (nStartLim > DL_MH_START_MAX)
           OR (tTempConfirm <= T#0S) OR (tOverloadConfirm <= T#0S) OR (tFreqConfirm <= T#0S)
           OR (tFreqWindow <= tFreqConfirm);
IF bCfgBad THEN
    bCfgLatch := TRUE;
END_IF
IF fbTrigReset.Q AND (NOT bCfgBad) THEN
    bCfgLatch := FALSE;              // 组态锁存解除（复位沿 + 组态已改对）/ config latch cleared
    uErrorId  := 16#0000_0000;       // 码位随解除归零 / code cleared with the latch
END_IF
IF bCfgLatch THEN
    uErrorId  := 16#0003_0532;       // 故障级：组态非法 / fault: illegal configuration
    bErrorInt := TRUE;               // R45 配对 / paired with the code
    eStateInt := E_DL_MotorAoiState.eFault;
END_IF

(*------------------------------------------------------------------------------
 * 段 5｜判据求值：信号闸（非有限只判不锁）+ 三判据 + 滚动窗计数
 *      Criteria evaluation with the non-finite signal gate
 *-----------------------------------------------------------------------------*)
bSigBad := (fWindingTemp <> fWindingTemp) OR ((fWindingTemp - fWindingTemp) <> (fWindingTemp - fWindingTemp))
           OR (ABS(fWindingTemp) >= DL_MH_FIN_LIM)
           OR (fCurrent <> fCurrent) OR ((fCurrent - fCurrent) <> (fCurrent - fCurrent))
           OR (ABS(fCurrent) >= DL_MH_FIN_LIM);

fCurrentRatio := 0.0;                                   // 比值缺省 0（除子由组态闸保证 > 0）[倍] / ratio default
IF NOT bSigBad THEN
    fCurrentRatio := fCurrent / fRatedCurrent;          // 除前已闸：fRatedCurrent > 0（段 4）/ divisor gated above [倍]
END_IF

bTempCond := (NOT bSigBad) AND (fWindingTemp > fTempLim);
bOvldCond := (NOT bSigBad) AND (fCurrentRatio > fOverloadRatio);

(* 滚动窗启动计数：窗满即清零并重新起算（自复位），计数饱和闸防溢出 *)
IF fbTrigStart.Q THEN
    IF nStartCnt < DL_MH_START_MAX THEN
        nStartCnt := nStartCnt + 1;                     // 启动计数推进 [次] / count up
    END_IF
END_IF
IF tonFreqWin.Q THEN
    nStartCnt := 0;                                     // 窗满清零（自复位窗每周期一次）/ window rollover resets the count
END_IF
bFreqCond := (nStartCnt >= nStartLim) AND (NOT bSigBad);

(* 三计时器门控：判据成立 AND 未锁存 AND 非组态故障（R99 挂状态量与判据量） *)
tonTemp(IN := bTempCond AND (NOT bTempLatch) AND (NOT bCfgLatch), PT := tTempConfirm);
tonOverload(IN := bOvldCond AND (NOT bOvldLatch) AND (NOT bCfgLatch), PT := tOverloadConfirm);
tonFreq(IN := bFreqCond AND (NOT bFreqLatch) AND (NOT bCfgLatch), PT := tFreqConfirm);

(*------------------------------------------------------------------------------
 * 段 6｜主状态机（红线 R6）：ENUM + CASE + ELSE 兜底
 *      Main state machine, phase dwell semantics only
 *-----------------------------------------------------------------------------*)
CASE eStateInt OF

    E_DL_MotorAoiState.eIdle:
        IF bEnable AND (NOT bCfgLatch) THEN
            eStateInt := E_DL_MotorAoiState.eMonitor;    // 使能且组态合法进监视 / enabled
        END_IF

    E_DL_MotorAoiState.eMonitor:
        IF (NOT bEnable) OR bCfgLatch THEN
            eStateInt := E_DL_MotorAoiState.eIdle;
        ELSIF bTempLatch OR bOvldLatch OR bFreqLatch THEN
            eStateInt := E_DL_MotorAoiState.eTripped;    // 任一确认即停机型驻留 / any cause trips
        END_IF

    E_DL_MotorAoiState.eTripped:
        (* 解除路径（R152 自证可达）：复位沿 AND 三类判据本拍均已消失 AND 组态合法 *)
        IF fbTrigReset.Q AND (NOT bTempCond) AND (NOT bOvldCond) AND (NOT bFreqCond)
           AND (NOT bCfgBad) THEN
            bTempLatch := FALSE;                         // 三类锁存同沿解除 / three latches cleared together
            bOvldLatch := FALSE;
            bFreqLatch := FALSE;
            uErrorId   := 16#0000_0000;
            eStateInt  := E_DL_MotorAoiState.eMonitor;
        ELSIF (NOT bEnable) OR bCfgLatch THEN
            eStateInt  := E_DL_MotorAoiState.eIdle;
        END_IF

    E_DL_MotorAoiState.eFault:
        IF fbTrigReset.Q AND (NOT bCfgBad) THEN
            bCfgLatch := FALSE;                          // 解除路径 / clear path
            uErrorId  := 16#0000_0000;
            eStateInt := E_DL_MotorAoiState.eIdle;
        END_IF

    ELSE
        (* 非法状态拦截 / illegal state interception *)
        eStateInt := E_DL_MotorAoiState.eFault;
        uErrorId  := 16#0003_0532;
        bErrorInt := TRUE;

END_CASE;

(*------------------------------------------------------------------------------
 * 段 7｜确认到期消化：三类各自独立锁存 + 独立码位（R190 归因唯一）
 *      Confirm expiry digestion: three independent latches with three distinct codes
 *-----------------------------------------------------------------------------*)
IF tonTemp.Q AND (NOT bTempLatch) THEN
    bTempLatch := TRUE;              // 过温锁存 / over-temperature latched
    uErrorId   := 16#0003_0533;      // 故障级：过温确认 / fault: over-temperature confirmed
    bErrorInt  := TRUE;              // R45 配对 / paired with the code
    eStateInt  := E_DL_MotorAoiState.eTripped;
END_IF
IF tonOverload.Q AND (NOT bOvldLatch) THEN
    bOvldLatch := TRUE;              // 过载锁存 / overload latched
    uErrorId   := 16#0003_0534;      // 故障级：过载确认 / fault: overload confirmed
    bErrorInt  := TRUE;              // R45 配对 / paired with the code
    eStateInt  := E_DL_MotorAoiState.eTripped;
END_IF
IF tonFreq.Q AND (NOT bFreqLatch) THEN
    bFreqLatch := TRUE;              // 启停频繁锁存 / frequent-start latched
    uErrorId   := 16#0003_0535;      // 故障级：启停频繁确认 / fault: frequent starts confirmed
    bErrorInt  := TRUE;              // R45 配对 / paired with the code
    eStateInt  := E_DL_MotorAoiState.eTripped;
END_IF

(*------------------------------------------------------------------------------
 * 段 8｜输出单一出口（范式 P-05）：健康出口取最严
 *      Single output exit with the strictest NE107 verdict
 *-----------------------------------------------------------------------------*)
bOverTemp  := bTempLatch;
bOverload  := bOvldLatch;
bFreqStart := bFreqLatch;
bTripReq   := bTempLatch OR bOvldLatch OR bFreqLatch;

IF (NOT bEnable) OR bCfgLatch THEN
    eHealth := E_DL_Ne107Status.eUnknown;                        // 未使能 / 组态故障：未知（禁降级为 Ok）
ELSIF bTempLatch OR bOvldLatch OR bFreqLatch THEN
    eHealth := E_DL_Ne107Status.eFailure;                        // 已确认：最严等级
ELSIF bTempCond OR bOvldCond OR bFreqCond THEN
    eHealth := E_DL_Ne107Status.eMaintenanceReq;                 // 确认中：维护级
ELSE
    eHealth := E_DL_Ne107Status.eOk;                             // 三类判据均未成立
END_IF

bError := bErrorInt OR bCfgLatch OR (eStateInt = E_DL_MotorAoiState.eTripped);
eState := eStateInt;
END_FUNCTION_BLOCK

(* ---- FB_DL_MotorPtcThermistProtect.st ---- *)
(*==============================================================================
 * 组件名称 (Component)  : FB_DL_MotorPtcThermistProtect
 * 溯源说明 (Provenance) : 道莅 clean-room 防御性实现（LBP 深化 + 国产手册需求线）
 * 所属子库 (Sublibrary) : DL_Device / MotorProtect
 * 当前版本 (Version)    : 1.0.0
 * 兼容性   (Platform)   : CODESYS 3.5 / TwinCAT 3 / 汇川 InoProShop；
 *                         纯 IEC 61131-3（第 3 版），仅用标准库 TON
 * 组件分类 (Category)   : 功能块（FUNCTION_BLOCK）· PTC 热敏电阻绕组保护
 * 功能一句话 (Summary)  : DIN 44081 判据的 PTC 三态保护：断线/短路/跳闸 + 确认延时。
 * 边界与安全 (Boundary) : ①断线判定优先于跳闸（先判阻值域再判确认）；
 *                         ②跳闸锁存仅 bReset 可清，且 bReset 仅在阻值回落
 *                           正常带（低于跳闸阈值）后有效（防复位振荡）；
 *                         ③滤波电阻一阶惯性，NaN/负值样本拒收保持旧值；
 *                         ④确认 TON 无条件周期刷新；
 *                         ⑤跳闸态短路回路的 bReset 无效（验收向量 ③）。
 * 错误码    : 16#0003_0378 断线（阻值不低于断线阈值）——故障级（持续态）
 *             16#0003_0379 短路（阻值不高于短路阈值）——故障级（持续态）
 *             16#0003_037A 跳闸确认（阻值进入跳闸域经延时确认）——故障级（锁存）
 * 码位总账  : 16#0003_0378 用 / 16#0003_0379 用 / 16#0003_037A 用
 * 修改记录  : v1.0.0 R26 初版
 *==============================================================================*)
FUNCTION_BLOCK FB_DL_MotorPtcThermistProtect
VAR_INPUT
    fThermRes     : LREAL; // PTC 热敏电阻实测阻值 [Ω] / Measured PTC resistance [Ω]
    bSensorOk     : BOOL;  // 传感器通道自诊断 OK / Sensor channel self-check OK
    fTripRes      : LREAL; // 跳闸阻值阈值 [Ω]，默认 3300 / Trip resistance threshold [Ω]
    fOpenRes      : LREAL; // 断线阻值阈值 [Ω]，默认 8000 / Open-circuit threshold [Ω]
    fShortRes     : LREAL; // 短路阻值阈值 [Ω]，默认 50 / Short-circuit threshold [Ω]
    tConfirmDelay : TIME;  // 跳闸确认延时 [ms] / Trip confirm delay [ms]
    bReset        : BOOL;  // 复位指令（回落正常带后有效）/ Reset command (valid only back in normal band)
END_VAR
VAR_OUTPUT
    bTrip        : BOOL; // 跳闸锁存输出，仅 bReset 可清 / Trip latch, cleared only by reset
    bWarn        : BOOL; // 预警：阻值进入预警带（0.75 倍跳闸阈）/ Warning: resistance in pre-trip band
    bSensorFault : BOOL; // 传感器故障（断线或短路或通道失效）/ Sensor fault (open, short or channel)
    fResFiltered : LREAL; // 一阶滤波阻值 [Ω] / First-order filtered resistance [Ω]
    eErr         : UDINT; // 本周期错误码，0=无错 / Error code this cycle, 0 = none
END_VAR
VAR CONSTANT
    cWarnRatio : LREAL := 0.75; // 预警带占跳闸阈比例 / Warning band ratio of trip threshold
    cIFilter   : LREAL := 0.2;  // 一阶滤波新样本权重 / Filter weight of new sample
END_VAR
VAR
    tonTrip  : TON;   // 跳闸确认定时器（无条件刷新）/ Trip confirm timer
    bResValid: BOOL;  // 本拍样本合法性 / Sample validity this cycle
    fResGuard: LREAL; // 本拍阻值守卫副本 / Cycle resistance guard copy
    bInTripDom: BOOL; // 阻值处于跳闸域（断线短路之间）/ Resistance in trip domain
END_VAR

// ---------- 参数与样本防御（守卫副本先行） ----------
fResGuard := fThermRes;
bResValid := bSensorOk AND (fResGuard >= 0.0) AND (fResGuard <= fOpenRes * 2.0);
IF fResGuard <> fResGuard THEN
    bResValid := FALSE;                       // NaN 拒收 / NaN rejected
END_IF

// ---------- 滤波：合法样本一阶更新，拒收保持旧值 ----------
IF bResValid THEN
    fResFiltered := fResFiltered + cIFilter * (fResGuard - fResFiltered); // 一阶惯性 / First-order lag
END_IF

// ---------- 无条件周期刷新：跳闸确认定时器 ----------
bInTripDom := bResValid AND (fResFiltered >= fTripRes) AND (fResFiltered < fOpenRes);
tonTrip(IN := bInTripDom, PT := tConfirmDelay);

// ---------- 断线判定（优先级最高） ----------
bSensorFault := FALSE;
eErr := 0;
IF NOT bSensorOk THEN
    bSensorFault := TRUE;                     // 通道自诊断失效 / Channel self-check failed
    eErr := 16#0003_0378;                     // 复用断线码（通道失效同域）/ Open code reused for channel fault
ELSIF bResValid AND (fResFiltered >= fOpenRes) THEN
    bSensorFault := TRUE;                     // 阻值达断线域 / Resistance in open domain
    eErr := 16#0003_0378;                     // 断线码 / Open-circuit code
ELSIF bResValid AND (fResFiltered <= fShortRes) THEN
    bSensorFault := TRUE;                     // 阻值达短路域 / Resistance in short domain
    eErr := 16#0003_0379;                     // 短路码 / Short-circuit code
END_IF

// ---------- 跳闸锁存：确认定时器到时置位，复位需回落正常带 ----------
IF tonTrip.Q THEN
    bTrip := TRUE;                            // 跳闸锁存置位 / Trip latch set
    eErr := 16#0003_037A;                     // 跳闸确认码 / Trip confirm code
END_IF

// ---------- 复位仲裁：阻值回落正常带（低于跳闸阈）后 bReset 才有效 ----------
IF bTrip THEN
    IF bResValid AND (fResFiltered < fTripRes) AND bReset THEN
        bTrip := FALSE;                       // 合法复位解除锁存 / Legal reset clears latch
        eErr  := 0;                           // 复位同拍清码 / Code cleared on reset
    ELSE
        eErr := 16#0003_037A;                 // 锁存态保持跳闸码（含短路态下复位被拒）/ Trip code held while latched
    END_IF
END_IF

// ---------- 预警带：介于 0.75 倍跳闸阈与跳闸阈之间 ----------
bWarn := bResValid AND (fResFiltered >= fTripRes * cWarnRatio) AND (fResFiltered < fTripRes);

END_FUNCTION_BLOCK

(* ---- FB_DL_MultiPumpRotationCtrl.st ---- *)
// FB_DL_MultiPumpRotationCtrl v1.0.0
(*==============================================================================
 * 功能描述: C4 多泵轮换均衡。2~4 台泵按累计运行小时数均衡轮换：领泵运行时间达
 *           tMinRun、小时差超 fBalThr 时经 eSwitch 两相切换（先停旧领泵，停机窗
 *           tMinStop 满窗后再启新领泵）；泵故障自动退出轮换池并告警，全池故障进
 *           eFault 锁存，bReset 上升沿唯一迁出。
 * 接口契约: 输入 bEnable/fDtSec/nPumpCount/aPumpFault/tMinRun/tMinStop/fBalThr/bReset；
 *           输出 abPumpRun/nLeadPump/nPoolCnt/eState/eCause/bError/nErrId。
 * 边界: ① 组态闸：nPumpCount 出 [2,4]、fDtSec<=0、tMinRun/tMinStop<=T#0S、fBalThr<0
 *           或任一浮点引脚 NaN → 故障锁存；② 泵槽位按常量 4 固定遍历，超组态槽位不参与；
 *           ③ 两枚 TON + 一枚 R_TRIG 段 0 无条件周期刷新；④ 零全局耦合。
 * 码表: 16#0007_0301 故障级总码（组态非法/全池故障/非法相位，锁存至 bReset 上升沿）；
 *       16#0007_0401 信息级：泵因故障退出轮换池（告警，每拍重算）。
 * 修订历史: 2026-11-23  v1.0.0  R74 首版
 *==============================================================================*)

TYPE E_DL_MprState :
(
    eIdle   := 0,     // 待机（未使能或全停）/ Idle, disabled or all stopped
    eRun    := 10,    // 领泵运行相 / Lead pump running
    eSwitch := 20,    // 切换过渡相（旧领泵已停，等待停机窗）/ Switching transition, old lead stopped
    eFault  := 90     // 故障锁存相（仅复位沿迁出）/ Fault latched, exit by reset edge only
);
END_TYPE

TYPE E_DL_MprCause :
(
    eNone         := 0,   // 无故障成因 / No cause
    eCfgIllegal   := 1,   // 组态非法 / Illegal configuration
    eAllPumpFault := 2,   // 轮换池全空（全部泵故障）/ Rotation pool empty, all pumps faulted
    ePhaseBad     := 3    // 非法相位兜底 / Illegal phase fallback
);
END_TYPE

FUNCTION_BLOCK FB_DL_MultiPumpRotationCtrl
VAR_INPUT
    bEnable    : BOOL := FALSE;            // 使能（FALSE 全停回待机）[-] / Enable, FALSE stops all
    fDtSec     : REAL := 0.010;            // 任务周期 [s]，域 > 0 / Task period [s], domain > 0
    nPumpCount : INT := 3;                 // 参与轮换泵数 [台]，域 [2,4] / Pump count in rotation, domain 2..4
    aPumpFault : ARRAY[1..4] OF BOOL := [FALSE, FALSE, FALSE, FALSE];   // 各泵故障反馈（TRUE 退出轮换池）[-] / Per-pump fault feedback
    tMinRun    : TIME := T#600S;           // 领泵最小运行时间，域 > T#0S [ms] / Minimum lead run time, domain > T#0S
    tMinStop   : TIME := T#60S;            // 被停泵最小停机时间，域 > T#0S [ms] / Minimum stop time, domain > T#0S
    fBalThr    : REAL := 1.0;              // 小时均衡切换阈值，域 >= 0 [h] / Hour balance threshold [h]
    bReset     : BOOL := FALSE;            // 复位，上升沿清故障锁存 [-] / Reset, rising edge clears fault
END_VAR
VAR_OUTPUT
    abPumpRun  : ARRAY[1..4] OF BOOL;      // 各泵启停指令（TRUE=运行）[-] / Per-pump run command
    nLeadPump  : INT := 0;                 // 当前领泵号（0=无领泵）[泵号] / Current lead pump index, 0 = none
    nPoolCnt   : INT := 0;                 // 当前轮换池泵数 [台] / Current pool size
    eState     : E_DL_MprState;            // 状态出口，段尾单点映射 / State outlet
    eCause     : E_DL_MprCause;            // 故障成因出口（归因唯一） / Fault cause outlet
    bError     : BOOL;                     // 故障锁存标志 [-] / Fault latch flag
    nErrId     : UDINT;                    // 事件码，0 = 无事件 / Event code, 0 = none
END_VAR
VAR
    _eState    : E_DL_MprState := E_DL_MprState.eIdle;     // 内部相位（CASE 唯一写入目标） / Internal phase
    _eCause    : E_DL_MprCause := E_DL_MprCause.eNone;     // 故障成因锁存量 / Latched cause
    rtReset    : R_TRIG;                    // 复位沿实例，段 0 无条件刷新 / Reset edge instance
    tonMinRun  : TON;                       // 领泵最小运行计时，段 0 无条件刷新 / Lead min-run timer
    tonMinStop : TON;                       // 停机窗计时（eSwitch 相独占），段 0 无条件刷新 / Stop window timer
    _a_fHours  : ARRAY[1..4] OF REAL := [0.0, 0.0, 0.0, 0.0];   // 各泵累计运行小时 [h] / Per-pump accumulated run hours
    _nLead     : INT := 0;                  // 内部领泵号（锁存量）[泵号] / Internal lead pump index
    _nCand     : INT := 0;                  // 切换候选泵号（eSwitch 入相时锁定）[泵号] / Candidate pump locked at switch entry
    _nPoolCnt  : INT := 0;                  // 轮换池泵数工作值 [台] / Pool size working value
    _bCfgBad   : BOOL;                      // 组态非法当拍量 [-] / Illegal configuration this scan
    _bFault    : BOOL;                      // 故障锁存位（锁存量） / Latched fault bit
    _uFault    : UDINT;                     // 故障码锁存（锁存量） / Latched fault code
    _uInfo     : UDINT;                     // 信息码，每拍重算 / Info code, recomputed each scan
    _bAnyOut   : BOOL;                      // 本拍有泵退出轮换池当拍量 [-] / A pump left the pool this scan
    _iLoop     : INT;                       // 泵槽位遍历游标 [槽位] / Pump slot loop cursor
    _fBest     : REAL;                      // 最小小时数搜索工作值 [h] / Min-hours search working value
    _bFound    : BOOL;                      // 候选命中标志 [-] / Candidate found flag
END_VAR

(* —— 段 0：定时器与沿实例无条件周期刷新（禁置于 IF/CASE 内） —— *)
rtReset(CLK := bReset);                                            // 复位沿，每拍必调 / Reset edge, called every scan
tonMinRun(IN := (_eState = E_DL_MprState.eRun) AND (NOT _bFault), PT := tMinRun);   // 领泵运行计时 / Lead run timer
tonMinStop(IN := (_eState = E_DL_MprState.eSwitch), PT := tMinStop);               // 停机窗计时（切换相独占）/ Stop window timer

(* —— 段 1：单拍量预清零（锁存量 _bFault/_uFault/_a_fHours/_nLead 不入清单） —— *)
_uInfo   := 16#0000_0000;                                          // 信息码每拍重算 / Info recomputed every scan
bError   := FALSE;                                                 // 故障标志每拍预清（置位处同拍回填） / Error flag preset
_bAnyOut := FALSE;                                                 // 退池事件标志预清 / Pool-exit flag preset
abPumpRun[1] := FALSE;                                             // 各泵指令每拍预清，运行相同拍回填 / Pump commands preset
abPumpRun[2] := FALSE;                                             // 各泵指令预清 / Pump commands preset
abPumpRun[3] := FALSE;                                             // 各泵指令预清 / Pump commands preset
abPumpRun[4] := FALSE;                                             // 各泵指令预清 / Pump commands preset
nLeadPump := 0;                                                    // 领泵号出口预清（eRun 相回填） / Lead outlet preset

(* —— 段 2：组态域闸（覆盖全部参与判据引脚） —— *)
_bCfgBad := (nPumpCount < 2) OR (nPumpCount > 4)                   // 泵数域闸 / Pump count domain gate
         OR (fDtSec <= 0.0) OR (fDtSec <> fDtSec)                  // 周期域与 NaN 闸 / Period domain and NaN gate
         OR (fBalThr < 0.0) OR (fBalThr <> fBalThr)                // 阈值域与 NaN 闸 / Threshold domain and NaN gate
         OR (tMinRun <= T#0S) OR (tMinStop <= T#0S);               // 时间域闸 / Time domain gates

(* —— 段 3：轮换池统计（常量 4 槽遍历，超组态槽位不参与，防越界） —— *)
_nPoolCnt := 0;                                                    // 池数清零重算 / Pool count recomputed
FOR _iLoop := 1 TO 4 DO                                             // 固定 4 槽遍历（上界常量无越界） / Fixed four-slot traversal
    IF (_iLoop <= nPumpCount) AND aPumpFault[_iLoop] THEN          // 组态内槽位且故障 / Faulted slot inside configuration
        _bAnyOut := TRUE;                                          // 退池事件 / Pool-exit event
    END_IF
    IF (_iLoop <= nPumpCount) AND (NOT aPumpFault[_iLoop]) THEN    // 组态内健康槽位计入池 / Healthy slot joins pool
        _nPoolCnt := _nPoolCnt + 1;                                // 池数递增 / Pool count increments
    END_IF
END_FOR

(* —— 段 4：故障锁存与解除（R45 配对；解除式全当拍量） —— *)
IF _bCfgBad THEN                                                   // 组态非法 / Illegal configuration
    _uFault := 16#0007_0301;                                       // 故障级总码 / Fault-level code
    _bFault := TRUE;
    bError  := TRUE;
    _eCause := E_DL_MprCause.eCfgIllegal;                          // 归因：组态非法 / Cause: illegal configuration
END_IF
IF bEnable AND (NOT _bFault) AND (_nPoolCnt = 0) THEN              // 全池故障 / Pool empty
    _uFault := 16#0007_0301;
    _bFault := TRUE;
    bError  := TRUE;
    _eCause := E_DL_MprCause.eAllPumpFault;                        // 归因：全池故障 / Cause: pool empty
END_IF
IF _bAnyOut AND (NOT _bFault) THEN                                 // 泵退池告警（信息级，不锁存） / Pool-exit warning
    _uInfo := 16#0007_0401;                                        // 信息级：泵退出轮换池 / Info: pump left pool
END_IF
IF rtReset.Q AND (NOT _bCfgBad) THEN                               // 解除沿（当拍量，无锁存因子） / Release edge
    _bFault := FALSE;                                              // 清故障锁存 / Clear fault latch
    _uFault := 16#0000_0000;                                       // 清故障码 / Clear fault code
    _eCause := E_DL_MprCause.eNone;                                // 清成因 / Clear cause
    IF _eState = E_DL_MprState.eFault THEN
        _eState := E_DL_MprState.eIdle;                            // 故障相唯一迁出路径 / Sole exit from fault phase
    END_IF
END_IF

(* —— 段 5：相位机（ENUM 全成员显式标签 + ELSE 兜底） —— *)
CASE _eState OF

E_DL_MprState.eIdle:
    IF (NOT _bFault) AND bEnable AND (_nPoolCnt > 0) THEN          // 出口 1：使能且池非空，选最小小时泵为领泵 / Enable with non-empty pool
        _fBest  := 1.0E30;                                         // 搜索初值（远大于可行小时数） / Search seed
        _bFound := FALSE;                                          // 命中标志清零 / Found flag cleared
        FOR _iLoop := 1 TO nPumpCount DO                           // 组态内槽位搜索 / Search inside configuration
            IF (NOT aPumpFault[_iLoop]) AND (_a_fHours[_iLoop] < _fBest) THEN   // 健康且小时更小 / Healthy and fewer hours
                _fBest  := _a_fHours[_iLoop];                      // 记录最小值 / Record minimum
                _nLead  := _iLoop;                                 // 记录候选领泵 / Record candidate lead
                _bFound := TRUE;                                   // 命中 / Found
            END_IF
        END_FOR
        IF _bFound THEN
            _eState := E_DL_MprState.eRun;                         // 进运行相 / Enter run phase
        END_IF
    ELSIF _bFault THEN                                             // 出口 2：故障锁存 / Fault latched
        _eState := E_DL_MprState.eFault;
    END_IF

E_DL_MprState.eRun:
    IF (NOT bEnable) THEN                                          // 出口 1：撤使能全停回待机 / Disable stops all
        _eState := E_DL_MprState.eIdle;
    ELSIF aPumpFault[_nLead] THEN                                  // 出口 2：领泵故障 → 立即停旧领泵进切换相（跳过运行窗，安全侧） / Lead fault, stop now
        _nCand := 0;                                               // 候选待重选 / Candidate to be reselected
        _eState := E_DL_MprState.eSwitch;
    ELSIF _bFault OR (_nPoolCnt = 0) THEN                          // 出口 3：锁存或池空 / Fault or pool empty
        _eState := E_DL_MprState.eFault;
    ELSE
        _a_fHours[_nLead] := _a_fHours[_nLead] + fDtSec / 3600.0;  // 领泵小时累计 [h] / Lead hours accumulate
        _fBest  := 1.0E30;                                         // 备用候选搜索初值 / Search seed
        _bFound := FALSE;                                          // 命中标志清零 / Found flag cleared
        FOR _iLoop := 1 TO nPumpCount DO                           // 搜索除领泵外最小小时候选 / Search candidate excluding lead
            IF (_iLoop <> _nLead) AND (NOT aPumpFault[_iLoop]) AND (_a_fHours[_iLoop] < _fBest) THEN
                _fBest  := _a_fHours[_iLoop];                      // 记录最小值 / Record minimum
                _nCand  := _iLoop;                                 // 记录候选 / Record candidate
                _bFound := TRUE;                                   // 命中 / Found
            END_IF
        END_FOR
        IF _bFound AND tonMinRun.Q AND ((_a_fHours[_nLead] - _a_fHours[_nCand]) > fBalThr) THEN  // 均衡切换判据（运行窗满 + 小时差超阈） / Balance criteria
            _eState := E_DL_MprState.eSwitch;                      // 进切换过渡相（旧领泵停） / Enter switch transition
        END_IF
    END_IF

E_DL_MprState.eSwitch:
    IF (NOT bEnable) THEN                                          // 出口 1：撤使能回待机 / Disable to idle
        _eState := E_DL_MprState.eIdle;
    ELSIF _bFault THEN                                             // 出口 2：故障锁存 / Fault latched
        _eState := E_DL_MprState.eFault;
    ELSE
        IF (_nCand < 1) OR (aPumpFault[_nCand]) THEN               // 候选未定或已故障 → 重选 / Candidate invalid, reselect
            _fBest  := 1.0E30;                                     // 搜索初值 / Search seed
            _bFound := FALSE;                                      // 命中标志清零 / Found flag cleared
            FOR _iLoop := 1 TO nPumpCount DO                       // 全池重选最小小时泵 / Reselection over the full pool
                IF (NOT aPumpFault[_iLoop]) AND (_a_fHours[_iLoop] < _fBest) THEN
                    _fBest  := _a_fHours[_iLoop];                  // 记录最小值 / Record minimum
                    _nCand  := _iLoop;                             // 记录候选 / Record candidate
                    _bFound := TRUE;                               // 命中 / Found
                END_IF
            END_FOR
            IF NOT _bFound THEN
                _nCand := 0;                                       // 池空，候选清零 / Pool empty, candidate cleared
            END_IF
        END_IF
        IF (_nCand >= 1) AND tonMinStop.Q THEN                     // 停机窗满且候选有效 → 启新领泵 / Stop window elapsed, start new lead
            _nLead  := _nCand;                                     // 领泵交接 / Lead handover
            _nCand  := 0;                                          // 候选清零 / Candidate cleared
            _eState := E_DL_MprState.eRun;                         // 回运行相 / Back to run phase
        END_IF
    END_IF

E_DL_MprState.eFault:
    ;                                                              // 故障相：仅段 4 复位沿可迁出 / Only the reset edge leaves this phase

ELSE
    _uFault := 16#0007_0301;                                       // 故障级：非法相位兜底 / Illegal-phase fallback
    _bFault := TRUE;
    bError  := TRUE;
    _eCause := E_DL_MprCause.ePhaseBad;                            // 归因：非法相位 / Cause: illegal phase
    _eState := E_DL_MprState.eFault;                               // 强拉故障相 / Force fault phase

END_CASE

(* —— 段 6：出口单点映射（名实同源；锁存码回放；故障相安全侧全停） —— *)
IF _eState = E_DL_MprState.eRun THEN                               // 仅运行相输出领泵指令 / Run phase drives lead only
    abPumpRun[_nLead] := TRUE;                                     // 领泵指令置位 / Lead command set
    nLeadPump := _nLead;                                           // 领泵号出口 / Lead outlet
END_IF
nPoolCnt := _nPoolCnt;                                             // 池数出口 / Pool size outlet
IF _bFault THEN
    nErrId := _uFault;                                             // 故障锁存码回放 / Replay latched fault code
ELSE
    nErrId := _uInfo;                                              // 信息码 / Info code
END_IF
bError := _bFault;                                                 // 故障标志与锁存同源（名实双出口） / Flag from latch
eState := _eState;                                                 // 状态出口 / State outlet
eCause := _eCause;                                                 // 成因出口 / Cause outlet

END_FUNCTION_BLOCK

(* ---- FB_DL_NtcChannelHealth.st ---- *)
(*==============================================================================
 * 组件名称 (Component)  : FB_DL_NtcChannelHealth
 * 所属子库 (Sublibrary) : DL_Device
 * 当前版本 (Version)    : 1.0.0
 * 兼容性 (Platform)     : CODESYS 3.5 / TwinCAT 3 / InoProShop（纯标准元素，零方言）
 * 功能描述 (Function)   : NTC 通道健康度 0~100 评分与预警。按评分周期对三维度打分：
 *                         上游故障（有故障即 0 分）、长期漂移（超限按「限值/实测」折算）、
 *                         窗口噪声（同法），按组态权重加权并分档 Good/Watch/Warn/Bad。
 *                         权重和不为 100 时回退默认 40/40/20 并报组态错（不停摆但必须报）；
 *                         温度非有限则本周期不计分（记 0 分会把健康通道判死）。不做温度
 *                         换算、不做断线检测本身（由上游掩码注入）。
 * 溯源 (Origin)         : 道莅 clean-room 防御性实现
 * 本文件内含 (Contains) : TYPE E_DL_HealthGrade / FUNCTION_BLOCK FB_DL_NtcChannelHealth
 * 依赖 (Depends)        : 无（仅 Standard.library 的 ABS / MIN）
 * 红线自检 (Redline)    : 无外部全局变量、无硬件地址直引 ｜ 全变量中英双语同行注释
 *                         两个限值判零防除零 ｜ 温度非有限只跳过本周期、不清健康度 ｜
 *                         评分周期定时器与沿实例无条件周期刷新 ｜ 枚举显式赋值 ｜ CASE 含 ELSE
 * 错误码表 (Codes)      : 16#0003_03B1 就绪（评分正常或本周期未到期）
 *                         16#0003_03B2 信息级 温度非有限，本周期不计分（健康度保持上次值）
 *                         16#0003_03B3 故障级 组态非法（权重和 ≠100 已回退默认、限值 ≤0）
 *                         16#0003_03B4 故障级 断线累计达 3 次（更换建议触发条件之一）
 *                         16#0003_03B5 预留：本版不发码（下一轮区间起点，禁止回填）
 * 修订历史 (Revision)   : 2026-11-17  v1.0.0  首版入库 · R28 · 阶段三批 2
 * 验收向量 (Acceptance) : 正向 无故障、漂移 0.2/2.0 ℃、噪声 0.01/0.5 ℃、权重 40/40/20 →
 *                         健康度 100、Good
 *                         反向 断线位置位且漂移 5 ℃（限 2.0）→ 健康度 ≤60 且 bReplaceReq=TRUE；
 *                         漂移限给 0 → 16#0003_03B3；温度给 NaN → 16#0003_03B2 且健康度保持
 *============================================================================*)

(*-----------------------------------------------------------------------------
 * 枚举: E_DL_HealthGrade（归属本功能块，同文件发布，全库唯一定义）
 *----------------------------------------------------------------------------*)
TYPE E_DL_HealthGrade :
(
    eGood  := 0,    // 良好：健康度 ≥80 / Good, health of 80 or above
    eWatch := 10,   // 关注：健康度 60~79 / Watch, health from 60 to 79
    eWarn  := 20,   // 预警：健康度 40~59 / Warn, health from 40 to 59
    eBad   := 30    // 差：健康度 <40，需更换 / Bad, health below 40, replacement required
);
END_TYPE

FUNCTION_BLOCK FB_DL_NtcChannelHealth
VAR_INPUT
    bEnable        : BOOL := FALSE;       // 使能 / Enable
    fTemp_C        : REAL := 25.0;        // 该通道温度 [℃] / Channel temperature in degrees Celsius
    uChFaultMask   : WORD;                // 上游通道故障掩码 [bit]，bit0 断线 bit1 短路 bit2 超域 / Upstream channel fault mask
    fDriftTotal_C  : REAL := 0.0;         // 长期漂移（对投运基线）[℃] / Long-term drift against the commissioning baseline
    fNoise_C       : REAL := 0.0;         // 窗口噪声（标准差）[℃] / Window noise as a standard deviation
    fDriftLimit_C  : REAL := 2.0;         // 漂移扣尽阈 [℃]，域 0.5~20 / Drift limit that zeroes the score, domain 0.5 to 20
    fNoiseLimit_C  : REAL := 0.5;         // 噪声扣尽阈 [℃]，域 0.05~5 / Noise limit that zeroes the score, domain 0.05 to 5
    uFaultWeight   : UINT := 40;          // 故障权重 [—]，域 0~100 / Fault weight, domain 0 to 100
    uDriftWeight   : UINT := 40;          // 漂移权重 [—]，域 0~100 / Drift weight, domain 0 to 100
    uNoiseWeight   : UINT := 20;          // 噪声权重 [—]，域 0~100 / Noise weight, domain 0 to 100
    tEvalPeriod    : TIME := T#5S;        // 评分周期 [ms]，域 1~60 s / Scoring period, domain 1 to 60 s
END_VAR
VAR_OUTPUT
    uHealth        : UINT := 100;         // 健康度 [0~100] / Health score from 0 to 100
    eGrade         : E_DL_HealthGrade;    // 健康分档 [—] / Health grade
    bReplaceReq    : BOOL;                // 更换建议（Bad 或断线累计 3 次） / Replacement advice
    bError         : BOOL;                // 故障级标志，仅故障级码置位 / Fault-class flag, set on fault codes only
    eErr           : UDINT;               // 错误码，段位 16#0003_xxxx / Error code in segment 16#0003_xxxx
END_VAR
VAR
    _bInit         : BOOL := FALSE;       // 首扫标志，取非判定 / First-scan flag, tested negated
    _bCfgOk        : BOOL;                // 组态合法标志 / Configuration valid flag
    _bFallback     : BOOL;                // 权重回退标志 / Weight fallback flag
    _bScoreNow     : BOOL;                // 本拍评分标志（周期到） / Score this scan flag
    _uwFault       : UINT := 40;          // 生效故障权重 / Effective fault weight
    _uwDrift       : UINT := 40;          // 生效漂移权重 / Effective drift weight
    _uwNoise       : UINT := 20;          // 生效噪声权重 / Effective noise weight
    _uwDisconnect  : UINT := 0;           // 断线累计次数 [次] / Disconnect count
    _uwFaultScore  : UINT;                // 故障维度得分 [0~100] / Fault dimension score
    _uwDriftScore  : UINT;                // 漂移维度得分 [0~100] / Drift dimension score
    _uwNoiseScore  : UINT;                // 噪声维度得分 [0~100] / Noise dimension score
    _uwSum         : UDINT;               // 加权和中间量 / Weighted sum intermediate
    _fDriftRatio   : REAL;                // 漂移占比（限值/实测） / Drift ratio, limit over measurement
    _fNoiseRatio   : REAL;                // 噪声占比（限值/实测） / Noise ratio, limit over measurement
    _rtrigFault    : R_TRIG;              // 断线位上升沿 / Rising edge of the disconnect bit
    _tonEval       : TON;                 // 评分周期计时（自复位） / Scoring period timer, self resetting
END_VAR
VAR CONSTANT
    DL_NTC_READY   : UDINT := 16#0003_03B1;  // 就绪码 / Ready code
    DL_NTC_SKIP    : UDINT := 16#0003_03B2;  // 信息级温度非有限码 / Info code for a non-finite temperature
    DL_NTC_CFG_BAD : UDINT := 16#0003_03B3;  // 故障级组态非法码 / Fault code for bad configuration
    DL_NTC_DISC    : UDINT := 16#0003_03B4;  // 故障级断线累计码 / Fault code for accumulated disconnections
    DL_NTC_BIT_DISC : WORD := 16#0001;       // 断线位 / Disconnect bit
    DL_NTC_DISC_MAX : UINT := 3;             // 断线累计阈值 [次] / Disconnect count threshold
    DL_NTC_DRIFT_LO : REAL := 0.5;           // 漂移限下限 [℃] / Drift limit lower bound
    DL_NTC_DRIFT_HI : REAL := 20.0;          // 漂移限上限 [℃] / Drift limit upper bound
    DL_NTC_NOISE_LO : REAL := 0.05;          // 噪声限下限 [℃] / Noise limit lower bound
    DL_NTC_NOISE_HI : REAL := 5.0;           // 噪声限上限 [℃] / Noise limit upper bound
    DL_NTC_GOOD     : UINT := 80;            // Good 档门限 / Good threshold
    DL_NTC_WATCH    : UINT := 60;            // Watch 档门限 / Watch threshold
    DL_NTC_WARN     : UINT := 40;            // Warn 档门限 / Warn threshold
    DL_NTC_HUNDRED  : REAL := 100.0;         // 百分比基准 / Percentage base
END_VAR

// 段 1｜输出与单拍标志预置
bError := FALSE;                                    // 故障标志预清 / Fault flag pre-cleared
eErr := 0;                                          // 错误码预清 / Error code pre-cleared
_bScoreNow := FALSE;                                // 评分标志预清 / Scoring flag pre-cleared

// 段 2｜沿检测与评分周期定时器无条件周期刷新（自复位：IN 取上一拍 Q 取非）
_rtrigFault(CLK := ((uChFaultMask AND DL_NTC_BIT_DISC) <> 16#0000));
_tonEval(IN := bEnable AND (NOT _tonEval.Q), PT := tEvalPeriod);
IF _tonEval.Q THEN
    _bScoreNow := TRUE;                             // 周期到：本拍评分 / The period elapsed, score this scan
END_IF

// 段 3｜首扫初始化（判据取非，R19）
IF NOT _bInit THEN
    uHealth := 100;                                 // 健康度起点 100 / Health starts at 100
    eGrade := E_DL_HealthGrade.eGood;               // 分档起点 Good / Grade starts good
    _bInit := TRUE;                                 // 首扫只做一次 / The first scan runs once
END_IF

// 段 4｜断线累计（上升沿计数，供更换建议）
IF _rtrigFault.Q THEN
    _uwDisconnect := _uwDisconnect + 1;             // 断线累计 +1 [次] / Disconnect count incremented
END_IF

// 段 5｜权重与限值组态闸（和 ≠100 → 回退 40/40/20 并报组态错；限值判零防除零）
_bFallback := (uFaultWeight + uDriftWeight + uNoiseWeight) <> 100;
IF _bFallback THEN
    _uwFault := 40;                                 // 回退故障权重 / Fallback fault weight
    _uwDrift := 40;                                 // 回退漂移权重 / Fallback drift weight
    _uwNoise := 20;                                 // 回退噪声权重 / Fallback noise weight
ELSE
    _uwFault := uFaultWeight;                       // 采用组态权重 / Use the configured weight
    _uwDrift := uDriftWeight;
    _uwNoise := uNoiseWeight;
END_IF
_bCfgOk := (NOT _bFallback)
        AND NOT ((fDriftLimit_C <> fDriftLimit_C) OR ((fDriftLimit_C - fDriftLimit_C) <> (fDriftLimit_C - fDriftLimit_C)))
        AND (fDriftLimit_C >= DL_NTC_DRIFT_LO) AND (fDriftLimit_C <= DL_NTC_DRIFT_HI)
        AND NOT ((fNoiseLimit_C <> fNoiseLimit_C) OR ((fNoiseLimit_C - fNoiseLimit_C) <> (fNoiseLimit_C - fNoiseLimit_C)))
        AND (fNoiseLimit_C >= DL_NTC_NOISE_LO) AND (fNoiseLimit_C <= DL_NTC_NOISE_HI)
        AND (tEvalPeriod >= T#1S) AND (tEvalPeriod <= T#60S);
IF NOT _bCfgOk THEN
    eErr := DL_NTC_CFG_BAD;                         // 故障级：组态非法 / Fault, bad configuration
    bError := TRUE;
END_IF
IF _uwDisconnect >= DL_NTC_DISC_MAX THEN
    eErr := DL_NTC_DISC;                            // 故障级：断线累计达阈值 / Fault, the disconnect count reached the threshold
    bError := TRUE;
END_IF

// 段 6｜评分（周期到且组态合法时才计分；温度非有限则本周期不计分）
IF _bScoreNow AND _bCfgOk THEN
    IF (fTemp_C <> fTemp_C) OR ((fTemp_C - fTemp_C) <> (fTemp_C - fTemp_C)) THEN
        eErr := DL_NTC_SKIP;                        // 信息级：温度非有限，本周期不计分 / Info, temperature not finite, no scoring this period
    ELSE
        // 故障维度：有任何上游故障位即 0 分
        IF uChFaultMask <> 16#0000 THEN
            _uwFaultScore := 0;                     // 故障维度 0 分 / Fault dimension scores zero
        ELSE
            _uwFaultScore := 100;                   // 故障维度满分 / Fault dimension scores full
        END_IF
        // 漂移维度：限内满分，超限按「限值 / 实测」折算
        IF ABS(fDriftTotal_C) <= fDriftLimit_C THEN
            _uwDriftScore := 100;
        ELSE
            _fDriftRatio := fDriftLimit_C / ABS(fDriftTotal_C);          // 占比 ≤1 / Ratio at most one
            _uwDriftScore := REAL_TO_UINT(_fDriftRatio * DL_NTC_HUNDRED);
        END_IF
        // 噪声维度：同法折算
        IF ABS(fNoise_C) <= fNoiseLimit_C THEN
            _uwNoiseScore := 100;
        ELSE
            _fNoiseRatio := fNoiseLimit_C / ABS(fNoise_C);               // 占比 ≤1 / Ratio at most one
            _uwNoiseScore := REAL_TO_UINT(_fNoiseRatio * DL_NTC_HUNDRED);
        END_IF
        // 加权合成（权重和恒为 100，除零不可达）
        _uwSum := (UINT_TO_UDINT(_uwFault) * UINT_TO_UDINT(_uwFaultScore)
                 + UINT_TO_UDINT(_uwDrift) * UINT_TO_UDINT(_uwDriftScore)
                 + UINT_TO_UDINT(_uwNoise) * UINT_TO_UDINT(_uwNoiseScore)) / 100;
        uHealth := UDINT_TO_UINT(_uwSum);           // 健康度落定 [0~100] / Health latched
    END_IF
END_IF

// 段 7｜分档（整数比较，禁浮点等判；ENUM + CASE + ELSE 兜底）
IF uHealth >= DL_NTC_GOOD THEN
    eGrade := E_DL_HealthGrade.eGood;
ELSIF uHealth >= DL_NTC_WATCH THEN
    eGrade := E_DL_HealthGrade.eWatch;
ELSIF uHealth >= DL_NTC_WARN THEN
    eGrade := E_DL_HealthGrade.eWarn;
ELSE
    eGrade := E_DL_HealthGrade.eBad;
END_IF
CASE eGrade OF
    E_DL_HealthGrade.eGood:
        bReplaceReq := FALSE;                       // Good 不建更换 / No replacement advice for good channels
    E_DL_HealthGrade.eWatch:
        bReplaceReq := FALSE;                       // Watch 暂不更换 / No replacement advice while watching
    E_DL_HealthGrade.eWarn:
        bReplaceReq := FALSE;                       // Warn 暂不更换 / No replacement advice while warning
    E_DL_HealthGrade.eBad:
        bReplaceReq := TRUE;                        // Bad 建议更换 / Replacement advised on bad channels
    ELSE
        // 非法分档兜底：按 Bad 处理（安全侧）并报组态错
        eGrade := E_DL_HealthGrade.eBad;
        bReplaceReq := TRUE;
        eErr := DL_NTC_CFG_BAD;                     // 故障级：分档非法 / Fault, illegal grade
        bError := TRUE;
END_CASE
IF (_uwDisconnect >= DL_NTC_DISC_MAX) THEN
    bReplaceReq := TRUE;                            // 断线累计达阈值亦建议更换 / Replacement also advised on repeated disconnections
END_IF
IF eErr = 0 THEN
    eErr := DL_NTC_READY;                           // 无事件回就绪码 / Ready code when nothing else applies
END_IF
END_FUNCTION_BLOCK

(* ---- FB_DL_OrificeDpZeroTrim.st ---- *)
(*
  FB_DL_OrificeDpZeroTrim  —  孔板差压零点漂移补偿 / Orifice DP zero-drift trim
  分类 Category : DL_Device
  码位 Code     : 16#03_2_1B
  段位说明      : 03_2 段低半字节已满，1x 段续号，1A 格由 CleaningBrushWear 启用，本件启用 1B 格（R192）
  版本 Version  : 1.0.0
  来源 Source   : t2-8-ne43 — 孔板计量零漂补偿待挖项
  溯源 Origin   : clean-room 实现，未复制任何源码行
                  （与 FC_DL_OrificeFlowCalc 分工：那件算流量，本件只供零点修正量，不算流量）
  功能 Function : 1) 静流时段判定：FC_DL_Deadband 归零型判 |fDpRawPa| 在静流带内 +
                  FB_DL_SignalStatistics 窗口峰峰值不超稳定阈（双判据防假静流）；
                  2) FB_DL_MedianFilter 对静流期样本取中值（抗单点毛刺），作为零漂观测值；
                  3) 静流持续 tZeroDwell（tonZero，单用途计时）→ 零点学习：
                  fZeroOffsetPa += (中值 − 旧零点) × fLearnRate（一阶趋近，学习率组态）；
                  4) 修正量出口：fDpCorrPa = fDpRawPa − fZeroOffsetPa（零点平移语义）。
  边界 Boundary : ① 本件只供修正量出口，不做流量换算、不做量程标定（分工见头注释）；
                  ② 零点学习值限幅 ±fTrimMaxPa（越限钳位 + 信息级码，防坏采样把零点学飞）；
                  ③ fLearnRate 域 (0, 1]，越域判组态故障（学习率 0 = 永不学习亦属组态错）；
                  ④ 非有限原始信号：保持上次有效值 + 信息级码（不中断，修正出口按保持值）；
                  ⑤ R228-A 达标声明：tonZero 单用途计时（IN = 静流判据电平），无跨相复用问题；
                  ⑥ R228-B 达标声明：eFault 迁出 = rtReset.Q（输入引脚，恒可达），逐字写于此。
  依赖 Depends  : FC_DL_Deadband（函数调用）；FB_DL_MedianFilter / FB_DL_SignalStatistics（实例化，引脚按 registry 实名）
  码表 Error codes（本件格 03_2_1B，子码步进 +0x100）:
    16#0003_011B 信息级：静流零点学习完成一次（本拍发生学习写入）
    16#0003_021B 故障级：组态非法（静流带/驻留时长/学习率/限幅域非法），锁存至复位
    16#0003_031B 故障级：保留码，本件无 CASE 主状态机，仅作后续维护者新增分支时的防御式默认码
    16#0003_041B 信息级：原始信号非有限，已保持上次有效值
    16#0003_051B 信息级：零点学习值越限幅，已钳制到 ±fTrimMaxPa

  修订历史 Revision :
    2026-11-19  v1.0.0  R39 首版（批次 3 · 序号 13）
*)

FUNCTION_BLOCK FB_DL_OrificeDpZeroTrim
VAR_INPUT
    fDpRawPa     : REAL := 0.0;       // 原始差压信号 [Pa] / Raw differential pressure signal
    fStaticBandPa: REAL := 20.0;      // 静流判定带半宽 [Pa]，域 > 0 / Static-flow band half width
    fStabRangePa : REAL := 10.0;      // 稳定判据峰峰值阈 [Pa]，域 > 0 / Stability peak-to-peak threshold
    tZeroDwell   : TIME := T#60S;     // 静流驻留学习时长 [ms]，域 > 0 / Static dwell before learning
    fLearnRate   : REAL := 0.2;       // 零点学习率 [无量纲 (0,1]] / Zero learning rate
    fTrimMaxPa   : REAL := 50.0;      // 零点学习值限幅 [Pa]，域 > 0 / Zero offset clamp
    nMedWindow   : INT  := 9;         // 中值窗长 [个]，3..15 奇数（越界钳位）/ Median window length
    bEnable      : BOOL := TRUE;      // 学习使能，FALSE 时只修正不学习 [-] / Learning enable
    bReset       : BOOL := FALSE;     // 故障复位，上升沿生效 / Fault reset, rising edge
    bZeroClr     : BOOL := FALSE;     // 零点清零沿，上升沿 fZeroOffsetPa 归零 / Zero offset clear, rising edge
END_VAR
VAR_OUTPUT
    fDpCorrPa    : REAL;              // 修正后差压 [Pa] = 原始 − 零点 / Corrected DP output
    fZeroOffsetPa: REAL;              // 当前零点学习值 [Pa] / Current learned zero offset
    bStaticFlow  : BOOL;              // 静流判定生效中 [-] / Static flow active flag
    bTrimValid   : BOOL;              // 修正有效（组态合法且输入有限）[-] / Trim validity flag
    bError       : BOOL;              // 故障锁存，仅故障级码置位，bReset 清除 [-] / Fault latch
    uErrorId     : UDINT;             // 事件码，0 = 无事件（故障级锁存回放）/ Event code
END_VAR
VAR
    fbMed      : FB_DL_MedianFilter;  // 中值滤波实例（主体首部无条件刷新）/ Median filter instance
    fbStat     : FB_DL_SignalStatistics;  // 差压统计窗实例（主体首部无条件刷新）/ DP statistics window instance
    tonZero    : TON;                 // 静流驻留计时（单用途，R228-A 口径）/ Static dwell timer, single purpose
    rtReset    : R_TRIG;              // 复位上升沿 / Reset rising edge
    rtZeroClr  : R_TRIG;              // 零点清零上升沿 / Zero clear rising edge
    _fDpEff    : REAL;                // 生效原始差压 [Pa]（非有限保持载体）/ Effective raw DP with hold carrier
    _fDpLast   : REAL := 0.0;         // 上次有效原始差压 [Pa] / Last valid raw DP
    _fZeroInt  : REAL := 0.0;         // 零点学习值内部量 [Pa]，出口镜像 / Internal zero offset register
    _bStaticDb : BOOL;                // 死区件静流判定 / Deadband static flag
    _bStatic   : BOOL;                // 双判据静流标志 / Combined static flag
    _bLearnEvt : BOOL;                // 本拍发生学习写入标志 / Learning write happened this cycle
    _bLearnBrk : BOOL;                // 学习拍断输入标志（TON 自复位纪律，用后即清）/ Learning break flag for timer reset
    _bRawBad   : BOOL;                // 本拍原始信号非有限标志 / Raw non-finite flag this cycle
    _uInfo     : UDINT;               // 信息码，每拍重算 / Info code
    _uFault    : UDINT;               // 故障码锁存寄存 / Latched fault code register
    _bFault    : BOOL;                // 故障锁存位 / Latched fault bit
    _bCfgBad   : BOOL;                // 组态非法聚合 / Configuration invalid aggregate
END_VAR
VAR CONSTANT
    DL_ODZ_INF_CAP : REAL := 1.0E15;  // 非有限值筛查幅值上限 / Non-finite screening cap
END_VAR

(* —— 段 0：定时器与边沿实例无条件周期刷新（R182：调用语句不得置于 IF/CASE 内） —— *)
rtReset(CLK := bReset);                                 // 复位沿刷新，每拍必调
rtZeroClr(CLK := bZeroClr);                             // 零点清零沿刷新，每拍必调
fbMed(fIn := _fDpEff,                                   // 中值滤波（输入为生效原始值）
      bSample := TRUE,                                  // 每拍采样（静流判据由外部承载）
      nWindow := nMedWindow,                            // 窗长（组态透传，内部钳位）
      bClear := FALSE);                                 // 不清窗（连续观测）
fbStat(fIn := _fDpEff,                                  // 统计窗（稳定判据用）
       bSample := TRUE,                                 // 每拍采样
       nWindow := 32,                                   // 窗长（稳定判据标准口径）
       bClear := FALSE);                                // 不清窗

(* —— 段 1：单拍量预清零（锁存量 _uFault/_bFault/_fZeroInt 不入清单，R187①） —— *)
_uInfo := 16#0000_0000;             // 信息码每拍重算
_bCfgBad := FALSE;                  // 组态非法预清零
_bLearnEvt := FALSE;                // 学习写入标志预清零
bStaticFlow := FALSE;               // 静流出口缺省 FALSE（段 4 单点重写）
uErrorId := 16#0000_0000;           // 事件码缺省无事件

(* —— 段 2：组态域闸（覆盖全部参与判据换算的引脚，R151；含除零口径） —— *)
IF (fStaticBandPa <= 0.0) OR (fStabRangePa <= 0.0) OR (fTrimMaxPa <= 0.0)
   OR (fLearnRate <= 0.0) OR (fLearnRate > 1.0)
   OR (TIME_TO_DINT(tZeroDwell) <= 0) THEN
    _bCfgBad := TRUE;               // 静流带/稳定阈/限幅/学习率/驻留域非法
END_IF

(* —— 段 3：故障锁存与迁出沿（R228-B：rtReset.Q 恒可达） —— *)
IF _bCfgBad AND (NOT _bFault) THEN
    _uFault := 16#0003_021B;        // 故障级：组态非法（仅首次进入时写入）
    _bFault := TRUE;
END_IF
IF rtReset.Q AND (NOT _bCfgBad) THEN
    _bFault := FALSE;               // 清故障锁存位（组态恢复合法为前提）
    _uFault := 16#0000_0000;
END_IF

(* —— 段 4：非有限防御与静流双判据 —— *)
_bRawBad := (fDpRawPa <> fDpRawPa) OR (ABS(fDpRawPa) > DL_ODZ_INF_CAP) OR ((fDpRawPa - fDpRawPa) <> 0.0);
IF _bRawBad THEN
    _fDpEff := _fDpLast;            // 非有限：保持上次有效值
    _uInfo := 16#0003_041B;         // 信息级：已保持
ELSE
    _fDpEff := fDpRawPa;            // 有效值入载体
    _fDpLast := fDpRawPa;
END_IF
_bStaticDb := (FC_DL_Deadband(fIn := _fDpEff,          // 归零型死区判静流带
                              fWidth := fStaticBandPa, // 带半宽
                              fCenter := 0.0,          // 零点中心
                              bZeroMode := TRUE) = 0.0);   // 归零型输出为 0 即在带内
IF (NOT _bRawBad) AND _bStaticDb AND fbStat.bValid AND (fbStat.fRange <= fStabRangePa) THEN
    _bStatic := TRUE;               // 双判据：带内 + 窗峰峰不超阈
ELSE
    _bStatic := FALSE;              // 任一判据不成立：非静流（TON 断输入即归零，R188）
END_IF
bStaticFlow := _bStatic;            // 静流出口镜像
tonZero(IN := _bStatic AND bEnable AND (NOT _bLearnBrk), PT := tZeroDwell);   // 静流驻留计时（顶层无条件调用；学习拍断输入一拍）
_bLearnBrk := FALSE;                // 断输入标志用后即清（R188 自复位纪律）

(* —— 段 5：零点学习（驻留到点 + 使能 + 组态合法） —— *)
IF tonZero.Q AND bEnable AND (NOT _bFault) THEN
    _fZeroInt := _fZeroInt + (fbMed.fMedian - _fZeroInt) * fLearnRate;   // 一阶趋近学习（中值抗毛刺）
    IF ABS(_fZeroInt) > fTrimMaxPa THEN
        _fZeroInt := MAX(-fTrimMaxPa, MIN(fTrimMaxPa, _fZeroInt));       // 限幅钳位
        _uInfo := 16#0003_051B;     // 信息级：学习值越限幅已钳制
    END_IF
    _bLearnEvt := TRUE;             // 本拍发生学习写入
    _bLearnBrk := TRUE;             // 学习拍断输入标志（下一拍复位驻留计时）
END_IF
IF rtZeroClr.Q THEN
    _fZeroInt := 0.0;               // 零点清零沿生效
END_IF
fZeroOffsetPa := _fZeroInt;         // 零点出口镜像
IF _bLearnEvt AND (NOT _bFault) THEN
    _uInfo := 16#0003_011B;         // 信息级：学习完成（覆盖限幅码优先级见两分支写入次序）
END_IF

(* —— 段 6：修正量出口（名实同源） —— *)
fDpCorrPa := _fDpEff - _fZeroInt;   // 修正 = 原始 − 零点（零点平移语义）
bTrimValid := (NOT _bFault) AND (NOT _bRawBad);   // 有效性 = 组态合法且输入有限

(* —— 段 7：事件码单点回放（故障锁存优先） —— *)
IF _bFault THEN
    uErrorId := _uFault;            // 故障锁存码回放
    bError := TRUE;
ELSE
    uErrorId := _uInfo;             // 信息码
    bError := FALSE;
END_IF

END_FUNCTION_BLOCK
